PROGRAM ModeManagement_モード管理
VAR
    Setting_M : BOOL;
    Manual_M : BOOL;
    Auto_M : BOOL;
    Dummy_M : BOOL;
    Inital_M : BOOL;
    Output_Error_M : ARRAY[0..99] OF Bool;
    Index_Error_001 : DINT;
    Index_B_001 : DINT;
    Index_Share_001 : DINT;
    Error_TON : ARRAY[0..99] OF TON;  (* [2] A(左側) ST1 測定タイムアウト; [4] A(左側) ST5 測定タイムアウト *)
    Error_TOF : ARRAY[0..99] OF TOF;
    AutoMode_A_M : ARRAY[0..99] OF Bool;
    ６ : DINT;
    ST4_A_Rev_01_Origin_M : ARRAY[0..99] OF Bool;  (* A(左側) ST4 反転1 原点復帰工程; [1] A(左側) ST4 反転1 原点復帰開始; [2] A(左側) ST4 反転1 原点復帰中; [3] A(左側) ST4 反転1 ピックアップ戻; [4] A(左側) ST4 反転1 モータ原点復帰開始; [5] A(左側) ST4 反転1 ピックアップ行; [6] A(左側) ST4 反転1 チャック閉; [7] A(左側) ST4 反転1 原点復帰完了（ワーク無） *)
    ST4_A_Rev_01_OriginDone : BOOL;  (* A(左側) ST4 反転1 原点復帰完了 *)
    ST4_A_Rev_02_Origin_M : ARRAY[0..99] OF Bool;  (* A(左側) ST6 反転2 原点復帰工程; [1] A(左側) ST6 反転2 原点復帰開始; [2] A(左側) ST6 反転2 原点復帰中; [3] A(左側) ST6 反転2 ピックアップ戻; [4] A(左側) ST6 反転2 モータ原点復帰開始; [5] A(左側) ST6 反転2 ピックアップ行; [6] A(左側) ST6 反転2 チャック閉; [7] A(左側) ST6 反転2 原点復帰完了（ワーク無） *)
    ST4_A_Rev_02_OriginDone : BOOL;  (* A(左側) ST6 反転2 原点復帰完了 *)
    ST4_B_Rev_01_Origin_M : ARRAY[0..99] OF Bool;  (* B(右側) ST4 反転1 原点復帰工程; [1] B(右側) ST4 反転1 原点復帰開始; [2] B(右側) ST4 反転1 原点復帰中; [3] B(右側) ST4 反転1 ピックアップ戻; [4] B(右側) ST4 反転1 モータ原点復帰開始; [5] B(右側) ST4 反転1 ピックアップ行; [6] B(右側) ST4 反転1 チャック閉; [7] B(右側) ST4 反転1 原点復帰完了（ワーク無） *)
    ST4_B_Rev_01_OriginDone : BOOL;  (* B(右側) ST4 反転1 原点復帰完了 *)
    ST4_B_Rev_02_Origin_M : ARRAY[0..99] OF Bool;  (* B(右側) ST6 反転2 原点復帰工程; [1] B(右側) ST6 反転2 原点復帰開始; [2] B(右側) ST6 反転2 原点復帰中; [3] B(右側) ST6 反転2 ピックアップ戻; [4] B(右側) ST6 反転2 モータ原点復帰開始; [5] B(右側) ST6 反転2 ピックアップ行; [6] B(右側) ST6 反転2 チャック閉; [7] B(右側) ST6 反転2 原点復帰完了（ワーク無） *)
    ST4_B_Rev_02_OriginDone : BOOL;  (* B(右側) ST6 反転2 原点復帰完了 *)
END_VAR
VAR_EXTERNAL
    Output_A_Error_M : ARRAY[0..99] OF Bool;
    Output_A_Restart_M : ARRAY[0..99] OF Bool;
    In_Sw_RESET : BOOL;
    In_Sw_START : BOOL;
    ManualMode : BOOL;
    M9999 : BOOL;
    Output_B_Error_M : ARRAY[0..99] OF Bool;  (* B(右側)シリンダエラー *)
    Output_B_Restart_M : ARRAY[0..99] OF Bool;  (* B(右側)シリンダ再開： *)
    Output_Share_Error_M : ARRAY[0..99] OF Bool;
    Output_Share_Restart_M : ARRAY[0..99] OF Bool;
    TimerQ_In_Sen_Accum_CV_A_Full : BOOL;
    Out_TDC_Stop : BOOL;
    In_Sen_Unl_Conv_A_Pass : BOOL;
    In_Sen_Accum_CV_A_Full : BOOL;
    In_Sen_Unl_Conv_B_Pass : BOOL;
    Pause : ARRAY[0..99] OF Bool;  (* [3] FH A(左側) ST1; [9] FH A(左側) ST5; [10] FH B(右側) ST1; [11] FH B(右側) ST5; [12] A(左側) ST6 反転2 ワーク不一致 *)
    AutoMode : BOOL;
    In_Sen_DOOR_01 : BOOL;
    In_Sen_DOOR_02 : BOOL;
    In_Sen_DOOR_03 : BOOL;
    In_Sen_DOOR_04 : BOOL;
    In_Sen_DOOR_05 : BOOL;
    In_Sen_DOOR_06 : BOOL;
    In_Sw_EMS1 : BOOL;
    In_Sw_EMS2 : BOOL;
    In_Sw_EMS3 : BOOL;
    In_Sen_AIR１_Pressure_01 : BOOL;
    In_Sen_AIR１_Pressure_02 : BOOL;
    In_Sen_AIR１_Pressure_03 : BOOL;
    TEST_M : ARRAY[0..99] OF Bool;
    ST0_Sup_Start : BOOL;  (* ST0_動作開始 *)
    Out_CYw_Sply_Pick_A_H_Auto : ARRAY[0..10] OF Bool;
    Out_CYw_Sply_Pick_A_H_Done : BOOL;
    Out_CYw_Sply_Slide_A_H_Auto : ARRAY[0..10] OF Bool;
    Out_CYw_Sply_Slide_A_H_Done : BOOL;
    Out_CYw_Sup_Chuck_A_Cl_H_Auto : ARRAY[0..10] OF Bool;
    Out_CYw_Sup_Chuck_A_Cl_H_Done : BOOL;
    In_Sen_Accum_CV_A_Arrival : BOOL;
    In_Sen_Work_A_Pos_00 : BOOL;
    Out_CYw_Sply_Pick_A_F_Auto : ARRAY[0..10] OF Bool;
    Out_CYw_Sply_Pick_A_F_Done : BOOL;
    Out_CYw_Sup_Chuck_A_Cl_F_Auto : ARRAY[0..10] OF Bool;
    Out_CYw_Sup_Chuck_A_Cl_F_Done : BOOL;
    Out_CYw_Sply_Slide_A_F_Auto : ARRAY[0..10] OF Bool;
    Out_CYw_Sply_Slide_A_F_Done : BOOL;
    Ins_A_Cv_Error : BOOL;
    Station_A_Data : ARRAY[0..8] OF sData;
    Ins_A_Cv_M : ARRAY[0..99] OF Bool;
    HMI_MessageNo : ARRAY[0..9] OF UINT;
    FH_5552_10_A_Auto : BOOL;
    In_Sen_Accum_CV_B_Full : BOOL;
    FH_Line3_Error_Status_1 : BOOL;
    FH_Line0_Error_Status_1 : BOOL;
    FH_Line1_Error_Status_1 : BOOL;
    FH_Line2_Error_Status_1 : BOOL;
    FH_Line0_Error_Clear_1 : BOOL;
    FH_Line1_Error_Clear_1 : BOOL;
    FH_Line2_Error_Clear_1 : BOOL;
    FH_Line3_Error_Clear_1 : BOOL;
    Ins_A_Next_Cycle : BOOL;
    OriginDone : BOOL;  (* 原点復帰完了 *)
    DummyDone : BOOL;  (* ダミーチェック完了 *)
    HMI_CurrentPage : STRING[256];
    Ins_A_End : BOOL;
    Auto_A_Start : BOOL;  (* 自動運転 開始 *)
    Auto_Ready : BOOL;  (* 自動運転可能 *)
    ST0_A_Sup_Busy : BOOL;
    ST1_A_Ca1_Busy : BOOL;
    RCON1_1_IN_Alarm : BOOL;  (* 軸異常 *)
    RCON1_1_IN_EmergencyStop : BOOL;  (* 非常停止状態（監視） *)
    RCON1_1_Error : BOOL;  (* 異常予備（未接続） *)
    RCON1_1_IN_HomeDone : BOOL;  (* 原点復帰完了 *)
    RCON1_1_Error_Clear : BOOL;  (* 解除予備（未接続） *)
    Error_M : ARRAY[0..99] OF Bool;  (* エラー：; [1] シリンダ; [2] コンベア＆ドアセンサ; [3] FH A(左側) ST1; [4] A(左側)検査コンベア ワーク不一致; [5] RCON1-1 異常; [9] FH A(左側) ST5; [10] FH B(右側) ST1; [11] FH B(右側) ST5; [12] A(左側) ST6 反転2 ワーク不一致 *)
    ST1_A_Ca1_M : ARRAY[0..99] OF Bool;  (* [6] A(左側) ST1 検査前ワーク不一致 *)
    ST2_A_Hgt_M : ARRAY[0..99] OF Bool;
    ST3_A_Dis1_M : ARRAY[0..99] OF Bool;
    HMI_Home_SW : BOOL;
    Origin_Busy : BOOL;  (* 原点復帰中 *)
    Out_CYw_Rev_01_Pick_A_H_Origin : ARRAY[0..10] OF Bool;  (* 原点復帰【Y710】A(左側)ST4 反転1ピックアップ戻： *)
    Out_CYw_Rev_01_Pick_A_H_Done : BOOL;  (* 【Y710】A(左側)ST4 反転1ピックアップ戻 動作完了 *)
    Stm_A_Rev_Axis000_Origin : BOOL;  (* A(左側) ST4 反転1 モータ原点復帰開始 *)
    Stm_A_Rev_Axis000_OriginDone : BOOL;  (* A(左側) ST4 反転1 モータ原点復帰完了 *)
    Out_CYw_Rev_01_Pick_A_F_Origin : ARRAY[0..99] OF Bool;  (* 原点復帰【Y711】A(左側)ST4 反転1ピックアップ行： *)
    Out_CYw_Rev_01_Pick_A_F_Done : BOOL;  (* 【Y711】A(左側)ST4 反転1ピックアップ行 動作完了 *)
    Out_CYw_Rev_01_Chk_A_H_Origin : ARRAY[0..99] OF Bool;  (* 原点復帰【Y708】A(左側)ST4 反転1チャック閉： *)
    Out_CYw_Rev_01_Chk_A_H_Done : BOOL;  (* 【Y708】A(左側)ST4 反転1チャック閉 動作完了 *)
    TimerQ_In_Sen_Work_A_Pos_04 : BOOL;
    Out_CYw_Rev_02_Pick_A_H_Origin : ARRAY[0..10] OF Bool;  (* 原点復帰 【Y714】A(左側)ST6 反転2ピックアップ戻 *)
    Out_CYw_Rev_02_Pick_A_H_Done : BOOL;  (* 【Y714】A(左側)ST6 反転2ピックアップ戻 動作完了 *)
    Stm_A_Rev_Axis001_Origin : BOOL;  (* A(左側) ST6 反転2 モータ原点復帰開始 *)
    Stm_A_Rev_Axis001_OriginDone : BOOL;  (* A(左側) ST6 反転2 モータ原点復帰完了 *)
    Out_CYw_Rev_02_Pick_A_F_Origin : ARRAY[0..99] OF Bool;  (* 原点復帰 【Y715】A(左側)ST6 反転2ピックアップ行 *)
    Out_CYw_Rev_02_Pick_A_F_Done : BOOL;  (* 【Y715】A(左側)ST6 反転2ピックアップ行 動作完了 *)
    Out_CYw_Rev_02_Chk_A_H_Origin : ARRAY[0..99] OF Bool;  (* 原点復帰 【Y712】A(左側)ST6 反転2チャック閉 戻 *)
    Out_CYw_Rev_02_Chk_A_H_Done : BOOL;  (* 【Y712】A(左側)ST6 反転2チャック閉 戻 動作完了 *)
    TimerQ_In_Sen_Work_A_Pos_06 : BOOL;  (* 【X208】A(左側)ワーク位置6 *)
    Auto_B_Start : BOOL;  (* B(右側)自動運転開始（後続処理未接続） *)
    Out_CYw_Rev_01_Pick_B_H_Origin : ARRAY[0..10] OF Bool;  (* 原点復帰 【Y810】B(右側)ST4 反転1ピックアップ戻 *)
    Out_CYw_Rev_01_Pick_B_H_Done : BOOL;  (* 【Y810】B(右側)ST4 反転1ピックアップ戻 動作完了 *)
    Stm_B_Rev_Axis002_Origin : BOOL;  (* B(右側) ST4 反転1 モータ原点復帰開始 *)
    Stm_B_Rev_Axis002_OriginDone : BOOL;  (* B(右側) ST4 反転1 モータ原点復帰完了 *)
    Out_CYw_Rev_01_Pick_B_F_Origin : ARRAY[0..99] OF Bool;  (* 原点復帰 【Y811】B(右側)ST4 反転1ピックアップ行 *)
    Out_CYw_Rev_01_Pick_B_F_Done : BOOL;  (* 【Y811】B(右側)ST4 反転1ピックアップ行 動作完了 *)
    Out_CYw_Rev_01_Chk_B_H_Origin : ARRAY[0..99] OF Bool;  (* 原点復帰 【Y808】B(右側)ST4 反転1チャック閉 戻 *)
    Out_CYw_Rev_01_Chk_B_H_Done : BOOL;  (* 【Y808】B(右側)ST4 反転1チャック閉 戻 動作完了 *)
    TimerQ_In_Sen_Work_B_Pos_04 : BOOL;  (* 【X406】B(右側)ワーク位置4 *)
    Out_CYw_Rev_02_Pick_B_H_Origin : ARRAY[0..10] OF Bool;  (* 原点復帰 【Y814】B(右側)ST6 反転2ピックアップ戻 *)
    Out_CYw_Rev_02_Pick_B_H_Done : BOOL;  (* 【Y814】B(右側)ST6 反転2ピックアップ戻 動作完了 *)
    Stm_B_Rev_Axis003_Origin : BOOL;  (* B(右側) ST6 反転2 モータ原点復帰開始 *)
    Stm_B_Rev_Axis003_OriginDone : BOOL;  (* B(右側) ST6 反転2 モータ原点復帰完了 *)
    Out_CYw_Rev_02_Pick_B_F_Origin : ARRAY[0..99] OF Bool;  (* 原点復帰 【Y815】B(右側)ST6 反転2ピックアップ行 *)
    Out_CYw_Rev_02_Pick_B_F_Done : BOOL;  (* 【Y815】B(右側)ST6 反転2ピックアップ行 動作完了 *)
    Out_CYw_Rev_02_Chk_B_H_Origin : ARRAY[0..99] OF Bool;  (* 原点復帰 【Y812】B(右側)ST6 反転2チャック閉 戻 *)
    Out_CYw_Rev_02_Chk_B_H_Done : BOOL;  (* 【Y812】B(右側)ST6 反転2チャック閉 戻 動作完了 *)
    TimerQ_In_Sen_Work_B_Pos_06 : BOOL;  (* 【X408】B(右側)ワーク位置6 *)
    ST4_A_Rev1_M : ARRAY[0..99] OF Bool;  (* [10] A(左側) ST4 ワーク不一致エラー; [12] 【Y708】A(左側) ST4 反転1チャック閉 *)
    ST5_A_Ca2_M : ARRAY[0..99] OF Bool;  (* A(左側) ST5 カメラ2工程; [1] A(左側) ST5 カメラ2検査開始; [2] 【Y724】A(左側) ST5 ストッパー戻; [3] A(左側) ST5 ワーク有無判定; [4] A(左側) ST5 ワーク有; [5] A(左側) ST5 ワーク無; [6] A(左側) ST5 検査前ワーク不一致; [7] A(左側) ST5 FH測定開始 *)
    FH_A_ST5_Auto : BOOL;  (* A(左側) ST5 FH自動測定 *)
END_VAR
VAR_EXTERNAL CONSTANT
    ST6_A_Rev2_M : ARRAY[0..99] OF Bool;  (* A(左側) ST6 反転2工程; [1] A(左側) ST6 反転2 動作開始; [2] A(左側) ST6 反転2 【Y714】ピックアップ戻; [3] A(左側) ST6 反転2 【Y725】位置6ストッパー戻; [4] A(左側) ST6 反転2 原点角度転送; [5] A(左側) ST6 反転2 原点位置移動開始; [6] A(左側) ST6 反転2 原点位置移動完了; [7] A(左側) ST6 反転2 ワーク有無判定; [8] A(左側) ST6 反転2 ワーク有・前工程OK; [9] A(左側) ST6 反転2 ワーク無・前工程NG; [10] A(左側) ST6 反転2 ワーク不一致エラー; [11] A(左側) ST6 反転2 【Y715】反転前ピックアップ行; [12] A(左側) ST6 反転2 【Y712】チャック閉; [13] A(左側) ST6 反転2 【Y714】反転前ピックアップ戻; [14] A(左側) ST6 反転2 反転角度転送; [15] A(左側) ST6 反転2 反転位置移動完了; [16] A(左側) ST6 反転2 【Y715】設置ピックアップ行; [17] A(左側) ST6 反転2 【Y713】チャック開; [18] A(左側) ST6 反転2 【Y714】設置ピックアップ戻 *)
END_VAR
VAR_EXTERNAL
    ST7_A_Dis2_M : ARRAY[0..99] OF Bool;  (* [9] ST7 A ワーク有; [10] ST3 A ワーク無; [11] ST7 排出前ワーク不一致エラー; [12] コンベア下降 位置転送; [13] コンベア下降 移動開始; [14] 排出チャック開 行; [15] セイフティ上昇 位置転送; [16] セイフティ上昇 移動開始; [17] NG / フォルダストック 仕分け IAI移動位置 判定; [18] ストックフォルダ位置; [19] カメラ2 キズNG位置; [20] カメラ2 姿NG位置; [21] 排出フォルダ送り行; [22] SF/NG2左右 移動開始; [23] SF/NG2上下 目標位置転送; [24] ストックフォルダ カウントup; [25] カメラ キズNG位置; [26] カメラ 姿NG位置; [27] SF/NG2上下 移動開始; [28] 排出チャック戻／ワーク解放; [29] SF/NG2上下 原点位置転送; [30] SF/NG2上下 原点移動開始; [31] SF/NG2左右 原点位置転送; [32] 排出フォルダ送り戻; [33] 排出フォルダ戻完了 *)
END_VAR
VAR
    _p1 : BOOL;
    _p2 : BOOL;
    _p3 : BOOL;
    _p4 : BOOL;
    _p5 : BOOL;
    _p6 : BOOL;
    _p7 : BOOL;
    _p8 : BOOL;
    _p9 : BOOL;
    _p10 : BOOL;
    _p11 : BOOL;
    _p12 : BOOL;
    _p13 : BOOL;
    _p14 : BOOL;
    _p15 : BOOL;
    _p16 : BOOL;
    _p17 : BOOL;
    _p18 : BOOL;
    _p19 : BOOL;
    _p20 : BOOL;
    _p21 : BOOL;
    _p22 : BOOL;
    _p23 : BOOL;
    _p24 : BOOL;
    _e25 : R_TRIG;
    _e26 : R_TRIG;
    _e27 : R_TRIG;
    _e28 : R_TRIG;
    _e29 : R_TRIG;
    _e30 : R_TRIG;
    _e31 : R_TRIG;
    _e32 : R_TRIG;
    _e33 : R_TRIG;
    _p34 : BOOL;
    _p35 : BOOL;
    _p36 : BOOL;
    _p37 : BOOL;
    _p38 : BOOL;
    _p39 : BOOL;
    _p40 : BOOL;
    _e41 : R_TRIG;
    _p42 : BOOL;
    _e43 : R_TRIG;
    _e44 : R_TRIG;
    _e45 : R_TRIG;
    _e46 : R_TRIG;
    _e47 : R_TRIG;
    _e48 : R_TRIG;
    _e49 : R_TRIG;
    _p50 : BOOL;
    _p51 : BOOL;
    _p52 : BOOL;
    _p53 : BOOL;
    _p54 : BOOL;
    _p55 : BOOL;
    _p56 : BOOL;
END_VAR

(* Section Initial_初期化処理: ladder, written here as Structured Text *)

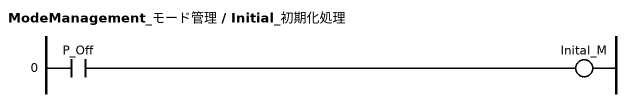
(* Rung 0 *)
Inital_M := P_Off;

(* Section Origin_原点復帰: ladder, written here as Structured Text *)

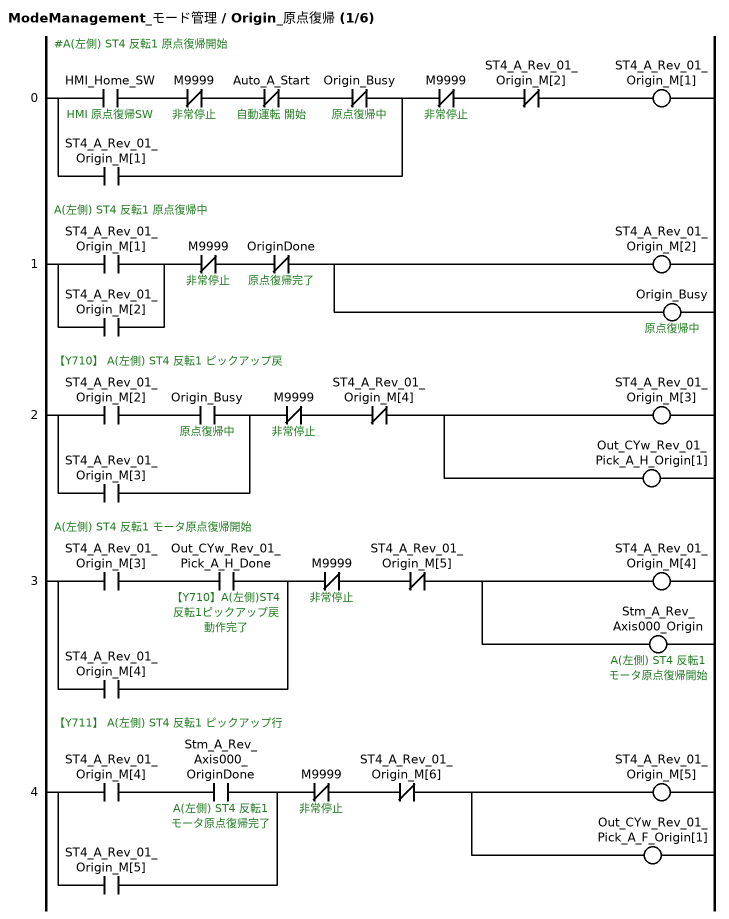
(* Rung 0: #A(左側) ST4 反転1 原点復帰開始 *)
ST4_A_Rev_01_Origin_M[1] := ((HMI_Home_SW AND NOT M9999 AND NOT Auto_A_Start AND NOT Origin_Busy) OR ST4_A_Rev_01_Origin_M[1]) AND NOT M9999 AND NOT ST4_A_Rev_01_Origin_M[2];
(* Rung 1: A(左側) ST4 反転1 原点復帰中 *)
_p1 := (ST4_A_Rev_01_Origin_M[1] OR ST4_A_Rev_01_Origin_M[2]) AND NOT M9999 AND NOT OriginDone;
ST4_A_Rev_01_Origin_M[2] := _p1;
Origin_Busy := _p1;
(* Rung 2: 【Y710】 A(左側) ST4 反転1 ピックアップ戻 *)
_p2 := ((ST4_A_Rev_01_Origin_M[2] AND Origin_Busy) OR ST4_A_Rev_01_Origin_M[3]) AND NOT M9999 AND NOT ST4_A_Rev_01_Origin_M[4];
ST4_A_Rev_01_Origin_M[3] := _p2;
Out_CYw_Rev_01_Pick_A_H_Origin[1] := _p2;
(* Rung 3: A(左側) ST4 反転1 モータ原点復帰開始 *)
_p3 := ((ST4_A_Rev_01_Origin_M[3] AND Out_CYw_Rev_01_Pick_A_H_Done) OR ST4_A_Rev_01_Origin_M[4]) AND NOT M9999 AND NOT ST4_A_Rev_01_Origin_M[5];
ST4_A_Rev_01_Origin_M[4] := _p3;
Stm_A_Rev_Axis000_Origin := _p3;
(* Rung 4: 【Y711】 A(左側) ST4 反転1 ピックアップ行 *)
_p4 := ((ST4_A_Rev_01_Origin_M[4] AND Stm_A_Rev_Axis000_OriginDone) OR ST4_A_Rev_01_Origin_M[5]) AND NOT M9999 AND NOT ST4_A_Rev_01_Origin_M[6];
ST4_A_Rev_01_Origin_M[5] := _p4;
Out_CYw_Rev_01_Pick_A_F_Origin[1] := _p4;

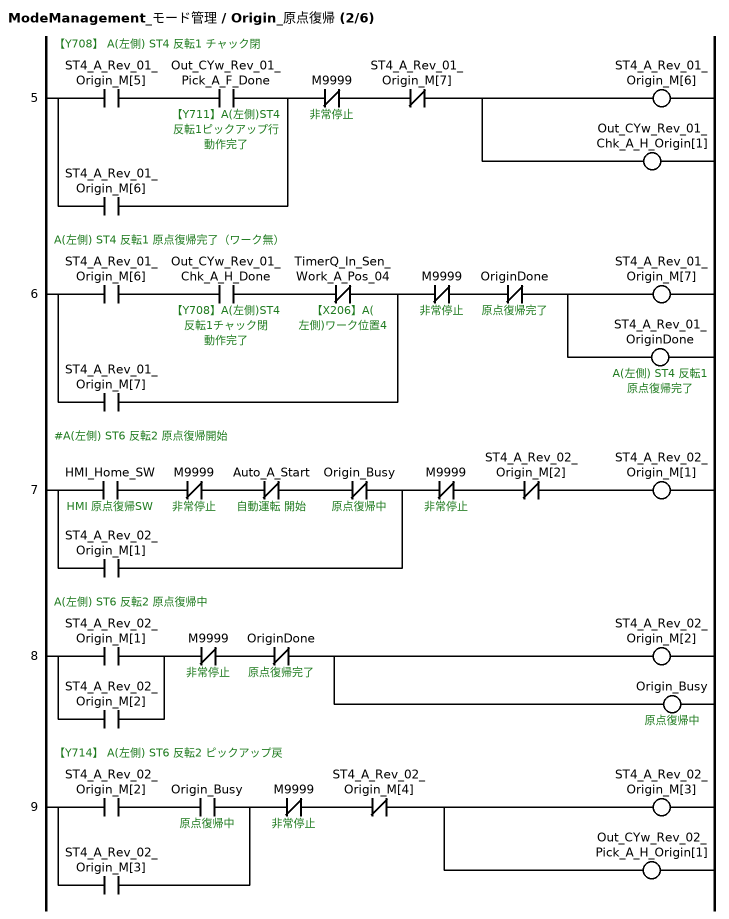
(* Rung 5: 【Y708】 A(左側) ST4 反転1 チャック閉 *)
_p5 := ((ST4_A_Rev_01_Origin_M[5] AND Out_CYw_Rev_01_Pick_A_F_Done) OR ST4_A_Rev_01_Origin_M[6]) AND NOT M9999 AND NOT ST4_A_Rev_01_Origin_M[7];
ST4_A_Rev_01_Origin_M[6] := _p5;
Out_CYw_Rev_01_Chk_A_H_Origin[1] := _p5;
(* Rung 6: A(左側) ST4 反転1 原点復帰完了（ワーク無） *)
_p6 := ((ST4_A_Rev_01_Origin_M[6] AND Out_CYw_Rev_01_Chk_A_H_Done AND NOT TimerQ_In_Sen_Work_A_Pos_04) OR ST4_A_Rev_01_Origin_M[7]) AND NOT M9999 AND NOT OriginDone;
ST4_A_Rev_01_Origin_M[7] := _p6;
ST4_A_Rev_01_OriginDone := _p6;
(* Rung 7: #A(左側) ST6 反転2 原点復帰開始 *)
ST4_A_Rev_02_Origin_M[1] := ((HMI_Home_SW AND NOT M9999 AND NOT Auto_A_Start AND NOT Origin_Busy) OR ST4_A_Rev_02_Origin_M[1]) AND NOT M9999 AND NOT ST4_A_Rev_02_Origin_M[2];
(* Rung 8: A(左側) ST6 反転2 原点復帰中 *)
_p7 := (ST4_A_Rev_02_Origin_M[1] OR ST4_A_Rev_02_Origin_M[2]) AND NOT M9999 AND NOT OriginDone;
ST4_A_Rev_02_Origin_M[2] := _p7;
Origin_Busy := _p7;
(* Rung 9: 【Y714】 A(左側) ST6 反転2 ピックアップ戻 *)
_p8 := ((ST4_A_Rev_02_Origin_M[2] AND Origin_Busy) OR ST4_A_Rev_02_Origin_M[3]) AND NOT M9999 AND NOT ST4_A_Rev_02_Origin_M[4];
ST4_A_Rev_02_Origin_M[3] := _p8;
Out_CYw_Rev_02_Pick_A_H_Origin[1] := _p8;

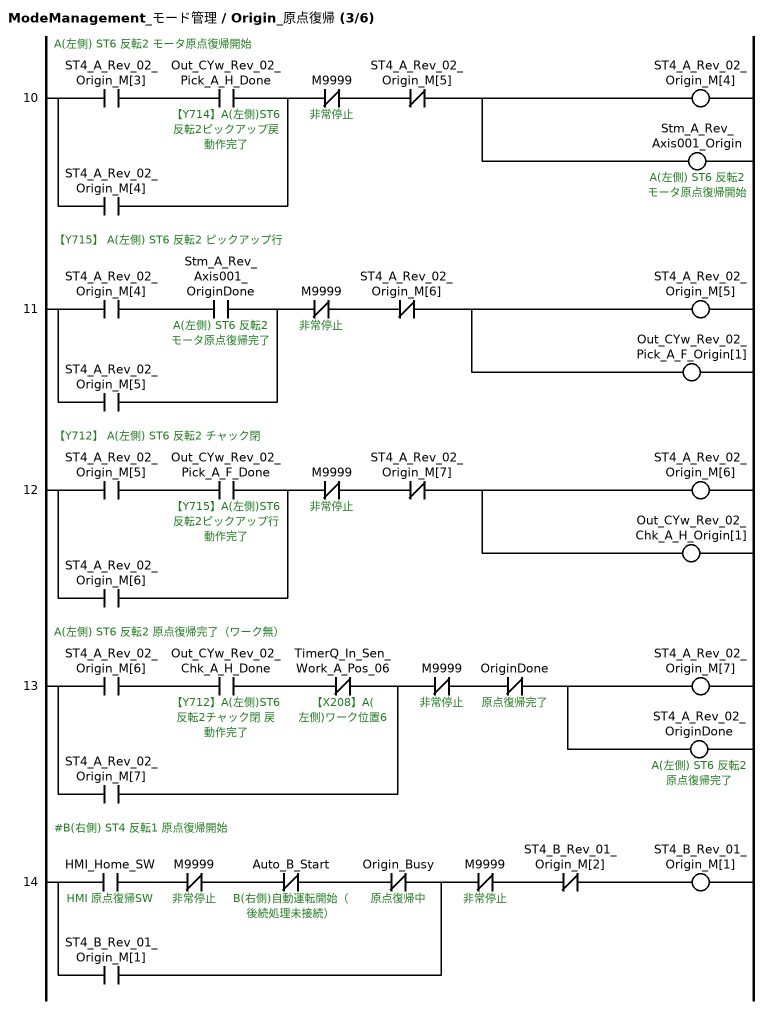
(* Rung 10: A(左側) ST6 反転2 モータ原点復帰開始 *)
_p9 := ((ST4_A_Rev_02_Origin_M[3] AND Out_CYw_Rev_02_Pick_A_H_Done) OR ST4_A_Rev_02_Origin_M[4]) AND NOT M9999 AND NOT ST4_A_Rev_02_Origin_M[5];
ST4_A_Rev_02_Origin_M[4] := _p9;
Stm_A_Rev_Axis001_Origin := _p9;
(* Rung 11: 【Y715】 A(左側) ST6 反転2 ピックアップ行 *)
_p10 := ((ST4_A_Rev_02_Origin_M[4] AND Stm_A_Rev_Axis001_OriginDone) OR ST4_A_Rev_02_Origin_M[5]) AND NOT M9999 AND NOT ST4_A_Rev_02_Origin_M[6];
ST4_A_Rev_02_Origin_M[5] := _p10;
Out_CYw_Rev_02_Pick_A_F_Origin[1] := _p10;
(* Rung 12: 【Y712】 A(左側) ST6 反転2 チャック閉 *)
_p11 := ((ST4_A_Rev_02_Origin_M[5] AND Out_CYw_Rev_02_Pick_A_F_Done) OR ST4_A_Rev_02_Origin_M[6]) AND NOT M9999 AND NOT ST4_A_Rev_02_Origin_M[7];
ST4_A_Rev_02_Origin_M[6] := _p11;
Out_CYw_Rev_02_Chk_A_H_Origin[1] := _p11;
(* Rung 13: A(左側) ST6 反転2 原点復帰完了（ワーク無） *)
_p12 := ((ST4_A_Rev_02_Origin_M[6] AND Out_CYw_Rev_02_Chk_A_H_Done AND NOT TimerQ_In_Sen_Work_A_Pos_06) OR ST4_A_Rev_02_Origin_M[7]) AND NOT M9999 AND NOT OriginDone;
ST4_A_Rev_02_Origin_M[7] := _p12;
ST4_A_Rev_02_OriginDone := _p12;
(* Rung 14: #B(右側) ST4 反転1 原点復帰開始 *)
ST4_B_Rev_01_Origin_M[1] := ((HMI_Home_SW AND NOT M9999 AND NOT Auto_B_Start AND NOT Origin_Busy) OR ST4_B_Rev_01_Origin_M[1]) AND NOT M9999 AND NOT ST4_B_Rev_01_Origin_M[2];

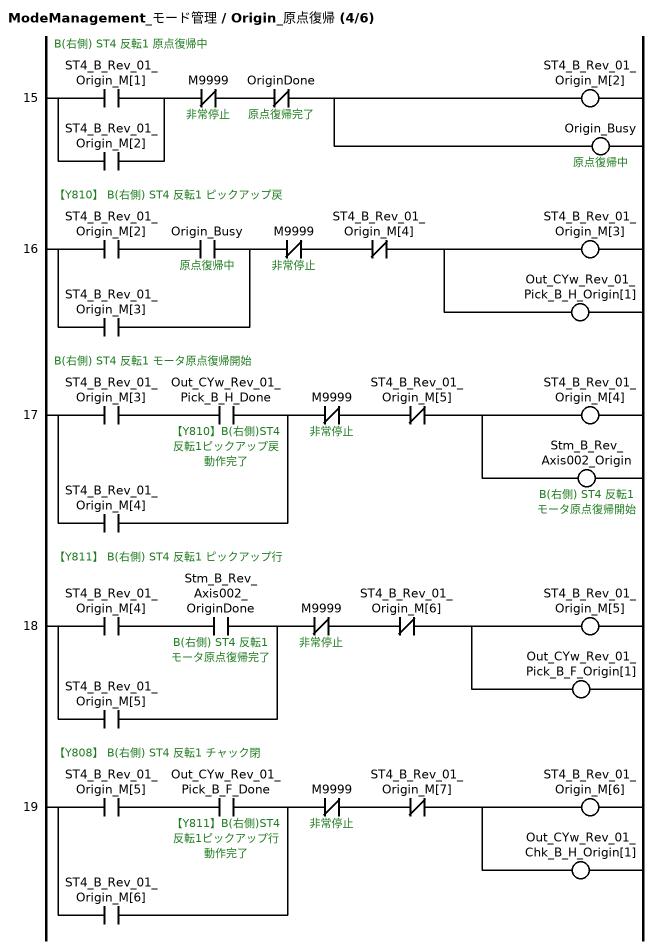
(* Rung 15: B(右側) ST4 反転1 原点復帰中 *)
_p13 := (ST4_B_Rev_01_Origin_M[1] OR ST4_B_Rev_01_Origin_M[2]) AND NOT M9999 AND NOT OriginDone;
ST4_B_Rev_01_Origin_M[2] := _p13;
Origin_Busy := _p13;
(* Rung 16: 【Y810】 B(右側) ST4 反転1 ピックアップ戻 *)
_p14 := ((ST4_B_Rev_01_Origin_M[2] AND Origin_Busy) OR ST4_B_Rev_01_Origin_M[3]) AND NOT M9999 AND NOT ST4_B_Rev_01_Origin_M[4];
ST4_B_Rev_01_Origin_M[3] := _p14;
Out_CYw_Rev_01_Pick_B_H_Origin[1] := _p14;
(* Rung 17: B(右側) ST4 反転1 モータ原点復帰開始 *)
_p15 := ((ST4_B_Rev_01_Origin_M[3] AND Out_CYw_Rev_01_Pick_B_H_Done) OR ST4_B_Rev_01_Origin_M[4]) AND NOT M9999 AND NOT ST4_B_Rev_01_Origin_M[5];
ST4_B_Rev_01_Origin_M[4] := _p15;
Stm_B_Rev_Axis002_Origin := _p15;
(* Rung 18: 【Y811】 B(右側) ST4 反転1 ピックアップ行 *)
_p16 := ((ST4_B_Rev_01_Origin_M[4] AND Stm_B_Rev_Axis002_OriginDone) OR ST4_B_Rev_01_Origin_M[5]) AND NOT M9999 AND NOT ST4_B_Rev_01_Origin_M[6];
ST4_B_Rev_01_Origin_M[5] := _p16;
Out_CYw_Rev_01_Pick_B_F_Origin[1] := _p16;
(* Rung 19: 【Y808】 B(右側) ST4 反転1 チャック閉 *)
_p17 := ((ST4_B_Rev_01_Origin_M[5] AND Out_CYw_Rev_01_Pick_B_F_Done) OR ST4_B_Rev_01_Origin_M[6]) AND NOT M9999 AND NOT ST4_B_Rev_01_Origin_M[7];
ST4_B_Rev_01_Origin_M[6] := _p17;
Out_CYw_Rev_01_Chk_B_H_Origin[1] := _p17;

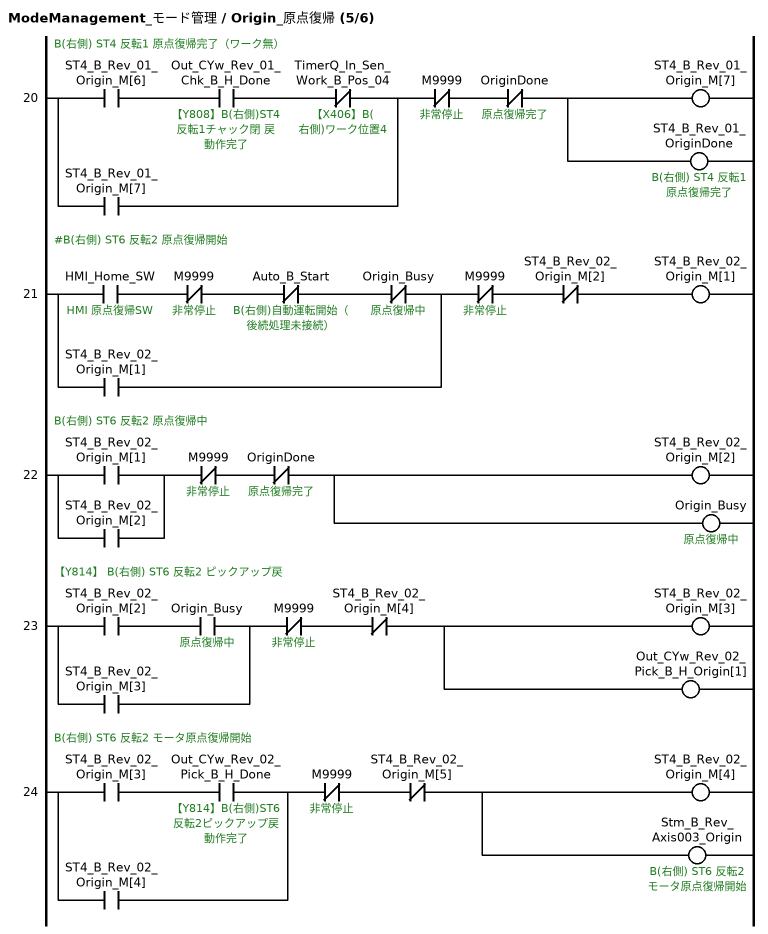
(* Rung 20: B(右側) ST4 反転1 原点復帰完了（ワーク無） *)
_p18 := ((ST4_B_Rev_01_Origin_M[6] AND Out_CYw_Rev_01_Chk_B_H_Done AND NOT TimerQ_In_Sen_Work_B_Pos_04) OR ST4_B_Rev_01_Origin_M[7]) AND NOT M9999 AND NOT OriginDone;
ST4_B_Rev_01_Origin_M[7] := _p18;
ST4_B_Rev_01_OriginDone := _p18;
(* Rung 21: #B(右側) ST6 反転2 原点復帰開始 *)
ST4_B_Rev_02_Origin_M[1] := ((HMI_Home_SW AND NOT M9999 AND NOT Auto_B_Start AND NOT Origin_Busy) OR ST4_B_Rev_02_Origin_M[1]) AND NOT M9999 AND NOT ST4_B_Rev_02_Origin_M[2];
(* Rung 22: B(右側) ST6 反転2 原点復帰中 *)
_p19 := (ST4_B_Rev_02_Origin_M[1] OR ST4_B_Rev_02_Origin_M[2]) AND NOT M9999 AND NOT OriginDone;
ST4_B_Rev_02_Origin_M[2] := _p19;
Origin_Busy := _p19;
(* Rung 23: 【Y814】 B(右側) ST6 反転2 ピックアップ戻 *)
_p20 := ((ST4_B_Rev_02_Origin_M[2] AND Origin_Busy) OR ST4_B_Rev_02_Origin_M[3]) AND NOT M9999 AND NOT ST4_B_Rev_02_Origin_M[4];
ST4_B_Rev_02_Origin_M[3] := _p20;
Out_CYw_Rev_02_Pick_B_H_Origin[1] := _p20;
(* Rung 24: B(右側) ST6 反転2 モータ原点復帰開始 *)
_p21 := ((ST4_B_Rev_02_Origin_M[3] AND Out_CYw_Rev_02_Pick_B_H_Done) OR ST4_B_Rev_02_Origin_M[4]) AND NOT M9999 AND NOT ST4_B_Rev_02_Origin_M[5];
ST4_B_Rev_02_Origin_M[4] := _p21;
Stm_B_Rev_Axis003_Origin := _p21;

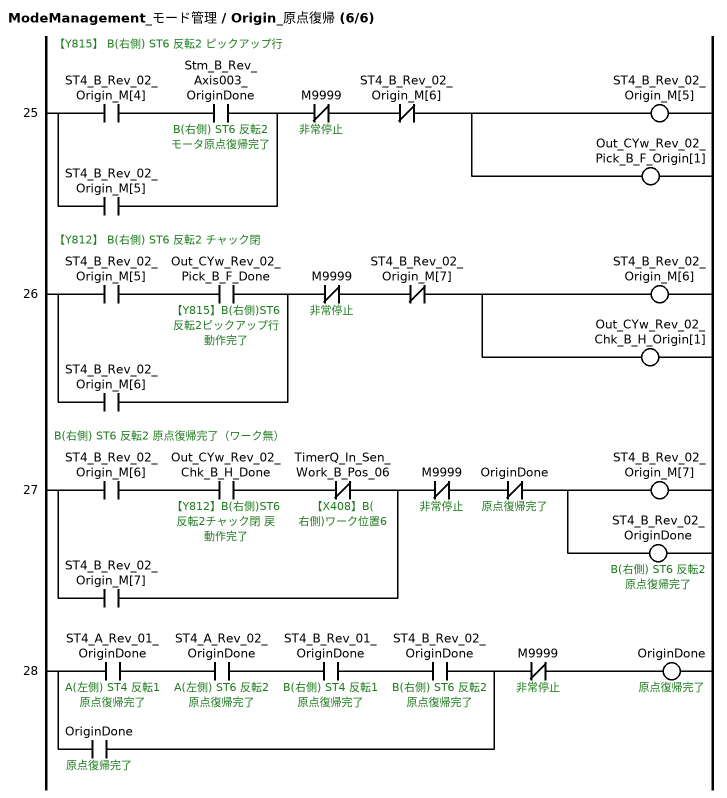
(* Rung 25: 【Y815】 B(右側) ST6 反転2 ピックアップ行 *)
_p22 := ((ST4_B_Rev_02_Origin_M[4] AND Stm_B_Rev_Axis003_OriginDone) OR ST4_B_Rev_02_Origin_M[5]) AND NOT M9999 AND NOT ST4_B_Rev_02_Origin_M[6];
ST4_B_Rev_02_Origin_M[5] := _p22;
Out_CYw_Rev_02_Pick_B_F_Origin[1] := _p22;
(* Rung 26: 【Y812】 B(右側) ST6 反転2 チャック閉 *)
_p23 := ((ST4_B_Rev_02_Origin_M[5] AND Out_CYw_Rev_02_Pick_B_F_Done) OR ST4_B_Rev_02_Origin_M[6]) AND NOT M9999 AND NOT ST4_B_Rev_02_Origin_M[7];
ST4_B_Rev_02_Origin_M[6] := _p23;
Out_CYw_Rev_02_Chk_B_H_Origin[1] := _p23;
(* Rung 27: B(右側) ST6 反転2 原点復帰完了（ワーク無） *)
_p24 := ((ST4_B_Rev_02_Origin_M[6] AND Out_CYw_Rev_02_Chk_B_H_Done AND NOT TimerQ_In_Sen_Work_B_Pos_06) OR ST4_B_Rev_02_Origin_M[7]) AND NOT M9999 AND NOT OriginDone;
ST4_B_Rev_02_Origin_M[7] := _p24;
ST4_B_Rev_02_OriginDone := _p24;
(* Rung 28 *)
OriginDone := ((ST4_A_Rev_01_OriginDone AND ST4_A_Rev_02_OriginDone AND ST4_B_Rev_01_OriginDone AND ST4_B_Rev_02_OriginDone) OR OriginDone) AND NOT M9999;

(* Section DummyCheck_ダミーチェック: ladder, written here as Structured Text *)

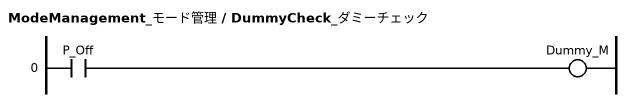
(* Rung 0 *)
Dummy_M := P_Off;

(* Section AutoMode_自動運転: ladder, written here as Structured Text *)

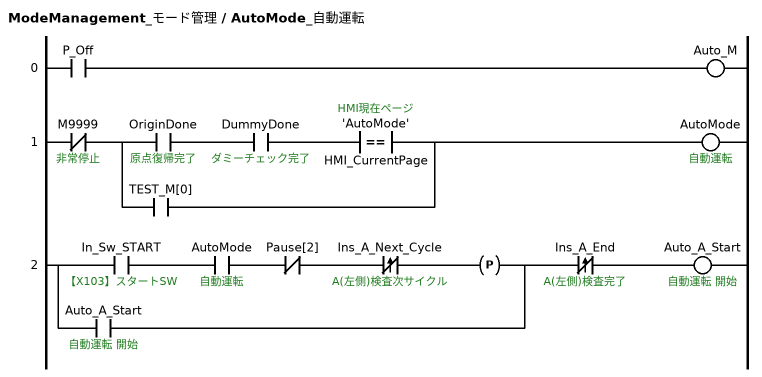
(* Rung 0 *)
Auto_M := P_Off;
(* Rung 1 *)
AutoMode := NOT M9999 AND ((OriginDone AND DummyDone AND ('AutoMode' = HMI_CurrentPage)) OR TEST_M[0]);
(* Rung 2 *)
_e25(CLK := Ins_A_Next_Cycle);
_e26(CLK := In_Sw_START AND AutoMode AND NOT Pause[2] AND NOT _e25.Q);
_e27(CLK := Ins_A_End);
Auto_A_Start := (_e26.Q OR Auto_A_Start) AND NOT _e27.Q;

(* Section Manual_手動運転: ladder, written here as Structured Text *)

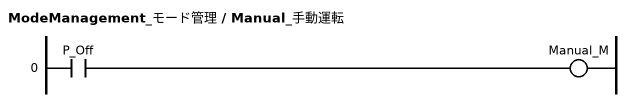
(* Rung 0 *)
Manual_M := P_Off;

(* Section Setting_設定: ladder, written here as Structured Text *)

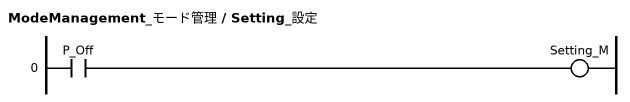
(* Rung 0 *)
Setting_M := P_Off;

(* Section Error_エラー処理: ladder, written here as Structured Text *)

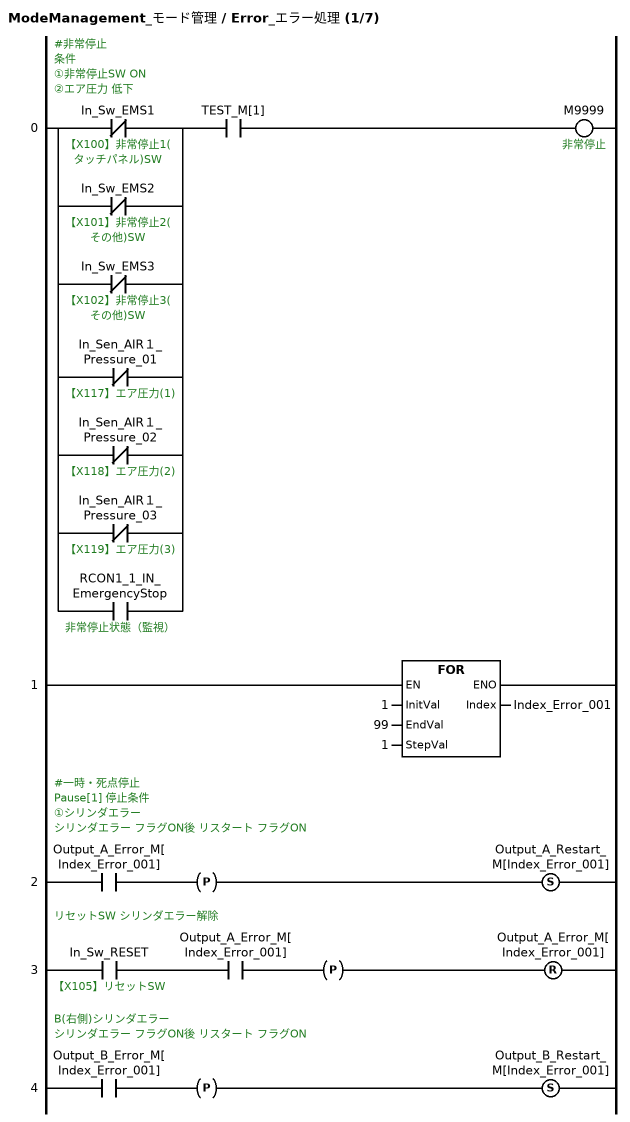
(* Rung 0: #非常停止 / 条件 / ①非常停止SW ON / ②エア圧力 低下 *)
M9999 := (NOT In_Sw_EMS1 OR NOT In_Sw_EMS2 OR NOT In_Sw_EMS3 OR NOT In_Sen_AIR１_Pressure_01 OR NOT In_Sen_AIR１_Pressure_02 OR NOT In_Sen_AIR１_Pressure_03 OR RCON1_1_IN_EmergencyStop) AND TEST_M[1];
(* Rung 1 *)
Index_Error_001 := FOR(InitVal := 1, EndVal := 99, StepVal := 1);
(* Rung 2: #一時・死点停止 / Pause[1] 停止条件 / ①シリンダエラー / シリンダエラー フラグON後 リスタート フラグON *)
_e28(CLK := Output_A_Error_M[Index_Error_001]);
IF _e28.Q THEN Output_A_Restart_M[Index_Error_001] := TRUE; END_IF;
(* Rung 3: リセットSW シリンダエラー解除 *)
_e29(CLK := In_Sw_RESET AND Output_A_Error_M[Index_Error_001]);
IF _e29.Q THEN Output_A_Error_M[Index_Error_001] := FALSE; END_IF;
(* Rung 4: B(右側)シリンダエラー / シリンダエラー フラグON後 リスタート フラグON *)
_e30(CLK := Output_B_Error_M[Index_Error_001]);
IF _e30.Q THEN Output_B_Restart_M[Index_Error_001] := TRUE; END_IF;

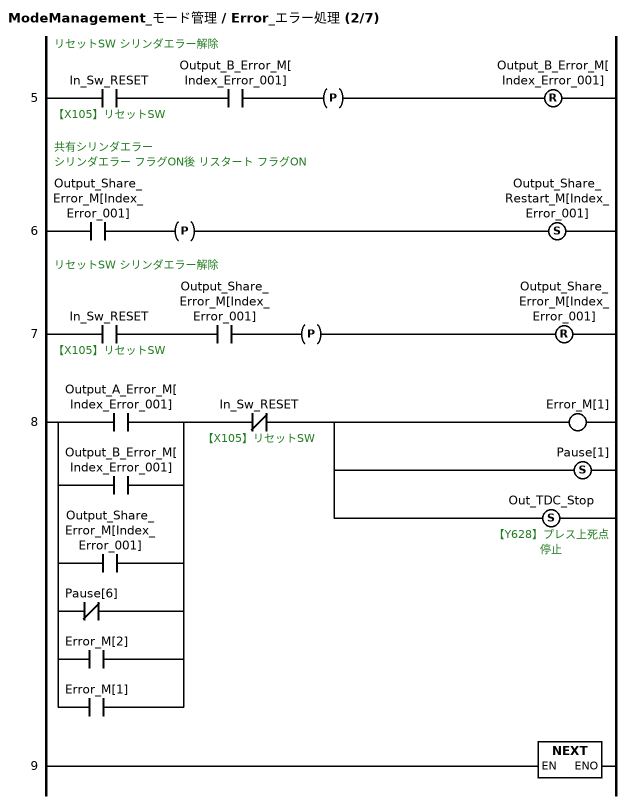
(* Rung 5: リセットSW シリンダエラー解除 *)
_e31(CLK := In_Sw_RESET AND Output_B_Error_M[Index_Error_001]);
IF _e31.Q THEN Output_B_Error_M[Index_Error_001] := FALSE; END_IF;
(* Rung 6: 共有シリンダエラー / シリンダエラー フラグON後 リスタート フラグON *)
_e32(CLK := Output_Share_Error_M[Index_Error_001]);
IF _e32.Q THEN Output_Share_Restart_M[Index_Error_001] := TRUE; END_IF;
(* Rung 7: リセットSW シリンダエラー解除 *)
_e33(CLK := In_Sw_RESET AND Output_Share_Error_M[Index_Error_001]);
IF _e33.Q THEN Output_Share_Error_M[Index_Error_001] := FALSE; END_IF;
(* Rung 8 *)
_p34 := (Output_A_Error_M[Index_Error_001] OR Output_B_Error_M[Index_Error_001] OR Output_Share_Error_M[Index_Error_001] OR NOT Pause[6] OR Error_M[2] OR Error_M[1]) AND NOT In_Sw_RESET;
Error_M[1] := _p34;
IF _p34 THEN
    Pause[1] := TRUE;
    Out_TDC_Stop := TRUE;
END_IF;
(* Rung 9 *)
NEXT();

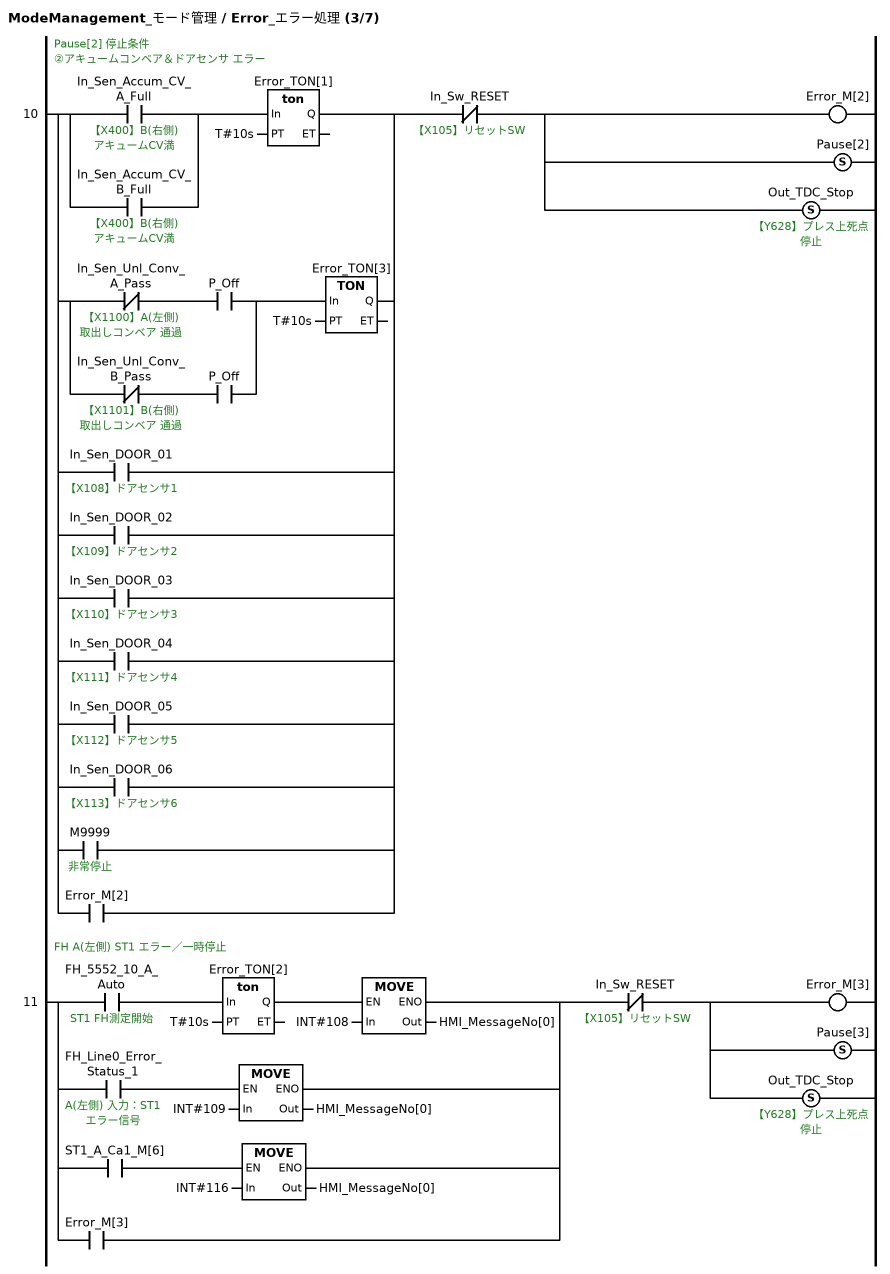
(* Rung 10: Pause[2] 停止条件 / ②アキュームコンベア＆ドアセンサ エラー *)
Error_TON[1](In := In_Sen_Accum_CV_A_Full OR In_Sen_Accum_CV_B_Full, PT := T#10s);
_p35 := Error_TON[1].Q;
Error_TON[3](In := (NOT In_Sen_Unl_Conv_A_Pass AND P_Off) OR (NOT In_Sen_Unl_Conv_B_Pass AND P_Off), PT := T#10s);
_p36 := (_p35 OR Error_TON[3].Q OR In_Sen_DOOR_01 OR In_Sen_DOOR_02 OR In_Sen_DOOR_03 OR In_Sen_DOOR_04 OR In_Sen_DOOR_05 OR In_Sen_DOOR_06 OR M9999 OR Error_M[2]) AND NOT In_Sw_RESET;
Error_M[2] := _p36;
IF _p36 THEN
    Pause[2] := TRUE;
    Out_TDC_Stop := TRUE;
END_IF;
(* Rung 11: FH A(左側) ST1 エラー／一時停止 *)
Error_TON[2](In := FH_5552_10_A_Auto, PT := T#10s);
IF Error_TON[2].Q THEN HMI_MessageNo[0] := INT#108; END_IF;
IF FH_Line0_Error_Status_1 THEN HMI_MessageNo[0] := INT#109; END_IF;
IF ST1_A_Ca1_M[6] THEN HMI_MessageNo[0] := INT#116; END_IF;
_p37 := (Error_TON[2].Q OR FH_Line0_Error_Status_1 OR ST1_A_Ca1_M[6] OR Error_M[3]) AND NOT In_Sw_RESET;
Error_M[3] := _p37;
IF _p37 THEN
    Pause[3] := TRUE;
    Out_TDC_Stop := TRUE;
END_IF;

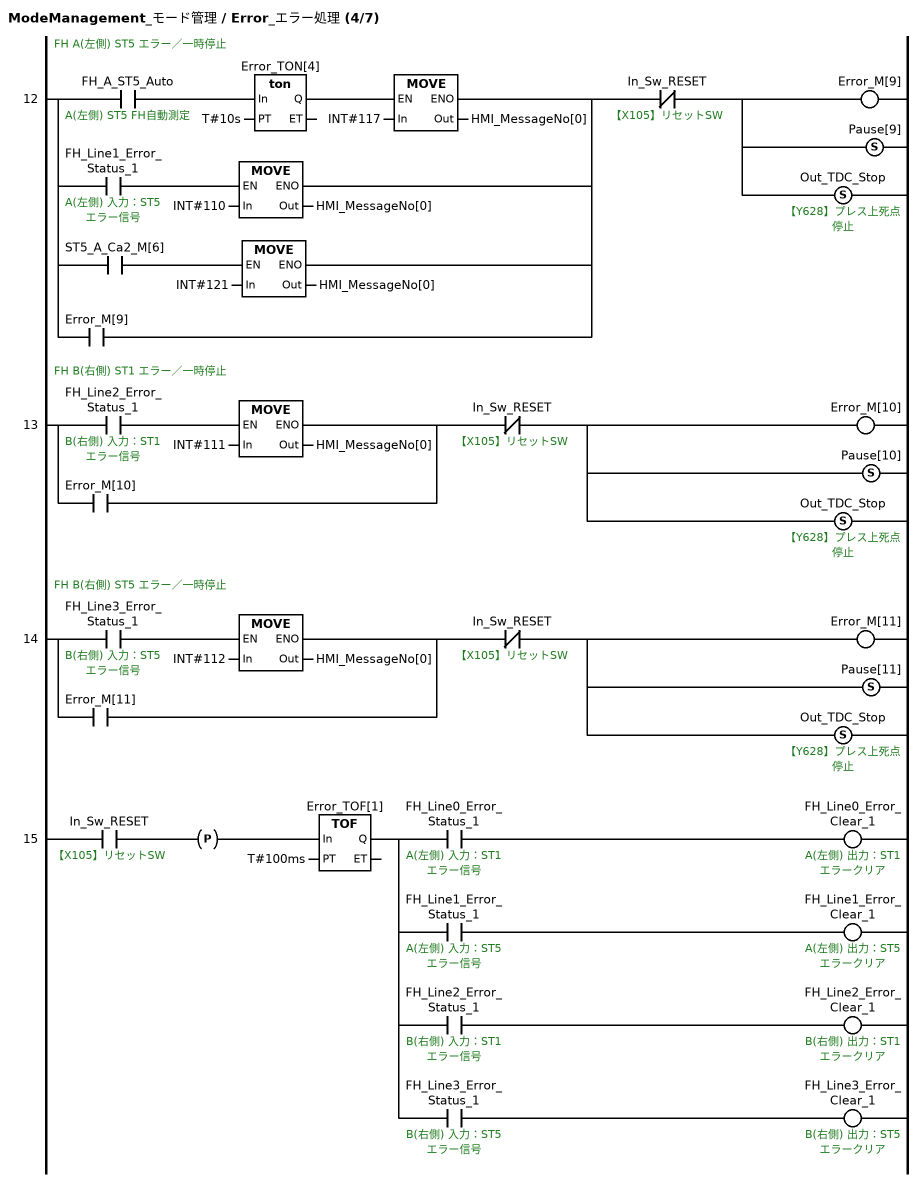
(* Rung 12: FH A(左側) ST5 エラー／一時停止 *)
Error_TON[4](In := FH_A_ST5_Auto, PT := T#10s);
IF Error_TON[4].Q THEN HMI_MessageNo[0] := INT#117; END_IF;
IF FH_Line1_Error_Status_1 THEN HMI_MessageNo[0] := INT#110; END_IF;
IF ST5_A_Ca2_M[6] THEN HMI_MessageNo[0] := INT#121; END_IF;
_p38 := (Error_TON[4].Q OR FH_Line1_Error_Status_1 OR ST5_A_Ca2_M[6] OR Error_M[9]) AND NOT In_Sw_RESET;
Error_M[9] := _p38;
IF _p38 THEN
    Pause[9] := TRUE;
    Out_TDC_Stop := TRUE;
END_IF;
(* Rung 13: FH B(右側) ST1 エラー／一時停止 *)
IF FH_Line2_Error_Status_1 THEN HMI_MessageNo[0] := INT#111; END_IF;
_p39 := (FH_Line2_Error_Status_1 OR Error_M[10]) AND NOT In_Sw_RESET;
Error_M[10] := _p39;
IF _p39 THEN
    Pause[10] := TRUE;
    Out_TDC_Stop := TRUE;
END_IF;
(* Rung 14: FH B(右側) ST5 エラー／一時停止 *)
IF FH_Line3_Error_Status_1 THEN HMI_MessageNo[0] := INT#112; END_IF;
_p40 := (FH_Line3_Error_Status_1 OR Error_M[11]) AND NOT In_Sw_RESET;
Error_M[11] := _p40;
IF _p40 THEN
    Pause[11] := TRUE;
    Out_TDC_Stop := TRUE;
END_IF;
(* Rung 15 *)
_e41(CLK := In_Sw_RESET);
Error_TOF[1](In := _e41.Q, PT := T#100ms);
FH_Line0_Error_Clear_1 := Error_TOF[1].Q AND FH_Line0_Error_Status_1;
FH_Line1_Error_Clear_1 := Error_TOF[1].Q AND FH_Line1_Error_Status_1;
FH_Line2_Error_Clear_1 := Error_TOF[1].Q AND FH_Line2_Error_Status_1;
FH_Line3_Error_Clear_1 := Error_TOF[1].Q AND FH_Line3_Error_Status_1;

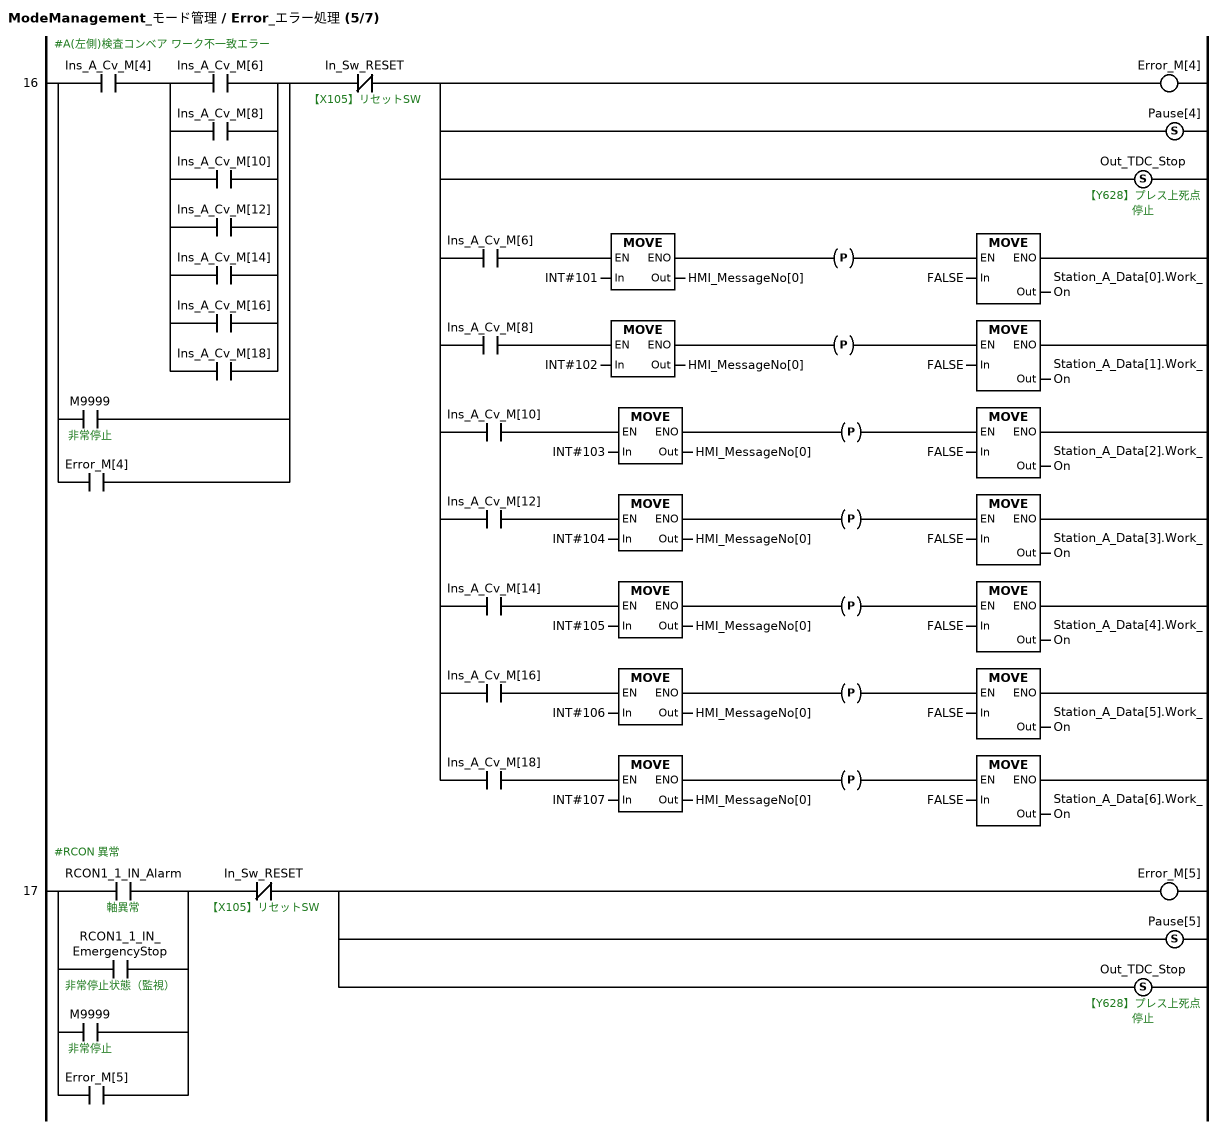
(* Rung 16: #A(左側)検査コンベア ワーク不一致エラー *)
_p42 := ((Ins_A_Cv_M[4] AND (Ins_A_Cv_M[6] OR Ins_A_Cv_M[8] OR Ins_A_Cv_M[10] OR Ins_A_Cv_M[12] OR Ins_A_Cv_M[14] OR Ins_A_Cv_M[16] OR Ins_A_Cv_M[18])) OR M9999 OR Error_M[4]) AND NOT In_Sw_RESET;
Error_M[4] := _p42;
IF _p42 THEN
    Pause[4] := TRUE;
    Out_TDC_Stop := TRUE;
END_IF;
IF _p42 AND Ins_A_Cv_M[6] THEN HMI_MessageNo[0] := INT#101; END_IF;
_e43(CLK := _p42 AND Ins_A_Cv_M[6]);
IF _e43.Q THEN Station_A_Data[0].Work_On := FALSE; END_IF;
IF _p42 AND Ins_A_Cv_M[8] THEN HMI_MessageNo[0] := INT#102; END_IF;
_e44(CLK := _p42 AND Ins_A_Cv_M[8]);
IF _e44.Q THEN Station_A_Data[1].Work_On := FALSE; END_IF;
IF _p42 AND Ins_A_Cv_M[10] THEN HMI_MessageNo[0] := INT#103; END_IF;
_e45(CLK := _p42 AND Ins_A_Cv_M[10]);
IF _e45.Q THEN Station_A_Data[2].Work_On := FALSE; END_IF;
IF _p42 AND Ins_A_Cv_M[12] THEN HMI_MessageNo[0] := INT#104; END_IF;
_e46(CLK := _p42 AND Ins_A_Cv_M[12]);
IF _e46.Q THEN Station_A_Data[3].Work_On := FALSE; END_IF;
IF _p42 AND Ins_A_Cv_M[14] THEN HMI_MessageNo[0] := INT#105; END_IF;
_e47(CLK := _p42 AND Ins_A_Cv_M[14]);
IF _e47.Q THEN Station_A_Data[4].Work_On := FALSE; END_IF;
IF _p42 AND Ins_A_Cv_M[16] THEN HMI_MessageNo[0] := INT#106; END_IF;
_e48(CLK := _p42 AND Ins_A_Cv_M[16]);
IF _e48.Q THEN Station_A_Data[5].Work_On := FALSE; END_IF;
IF _p42 AND Ins_A_Cv_M[18] THEN HMI_MessageNo[0] := INT#107; END_IF;
_e49(CLK := _p42 AND Ins_A_Cv_M[18]);
IF _e49.Q THEN Station_A_Data[6].Work_On := FALSE; END_IF;
(* Rung 17: #RCON 異常 *)
_p50 := (RCON1_1_IN_Alarm OR RCON1_1_IN_EmergencyStop OR M9999 OR Error_M[5]) AND NOT In_Sw_RESET;
Error_M[5] := _p50;
IF _p50 THEN
    Pause[5] := TRUE;
    Out_TDC_Stop := TRUE;
END_IF;

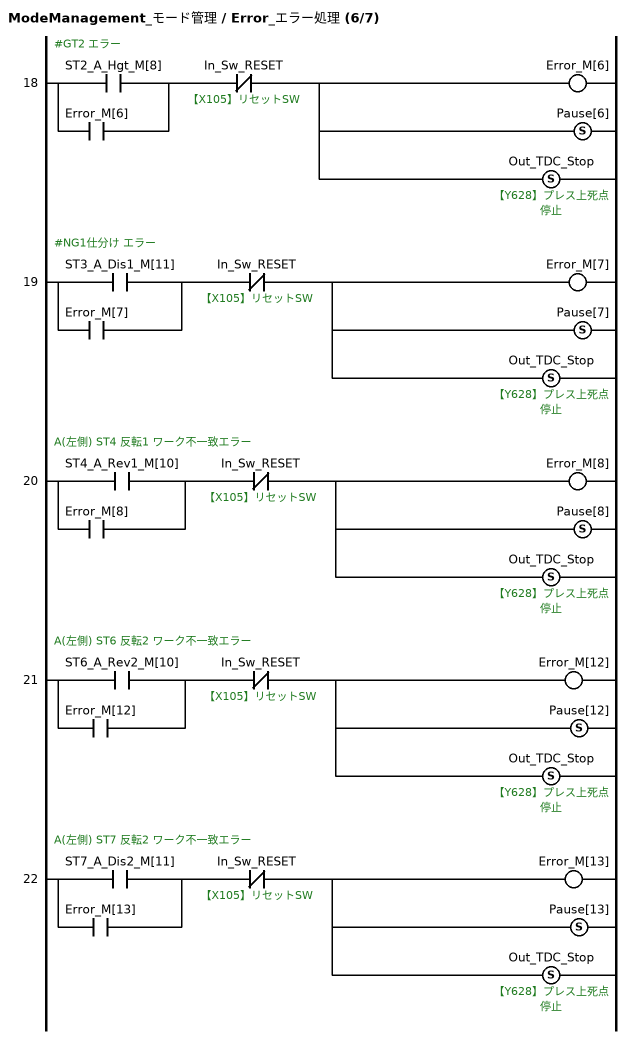
(* Rung 18: #GT2 エラー *)
_p51 := (ST2_A_Hgt_M[8] OR Error_M[6]) AND NOT In_Sw_RESET;
Error_M[6] := _p51;
IF _p51 THEN
    Pause[6] := TRUE;
    Out_TDC_Stop := TRUE;
END_IF;
(* Rung 19: #NG1仕分け エラー *)
_p52 := (ST3_A_Dis1_M[11] OR Error_M[7]) AND NOT In_Sw_RESET;
Error_M[7] := _p52;
IF _p52 THEN
    Pause[7] := TRUE;
    Out_TDC_Stop := TRUE;
END_IF;
(* Rung 20: A(左側) ST4 反転1 ワーク不一致エラー *)
_p53 := (ST4_A_Rev1_M[10] OR Error_M[8]) AND NOT In_Sw_RESET;
Error_M[8] := _p53;
IF _p53 THEN
    Pause[8] := TRUE;
    Out_TDC_Stop := TRUE;
END_IF;
(* Rung 21: A(左側) ST6 反転2 ワーク不一致エラー *)
_p54 := (ST6_A_Rev2_M[10] OR Error_M[12]) AND NOT In_Sw_RESET;
Error_M[12] := _p54;
IF _p54 THEN
    Pause[12] := TRUE;
    Out_TDC_Stop := TRUE;
END_IF;
(* Rung 22: A(左側) ST7 反転2 ワーク不一致エラー *)
_p55 := (ST7_A_Dis2_M[11] OR Error_M[13]) AND NOT In_Sw_RESET;
Error_M[13] := _p55;
IF _p55 THEN
    Pause[13] := TRUE;
    Out_TDC_Stop := TRUE;
END_IF;

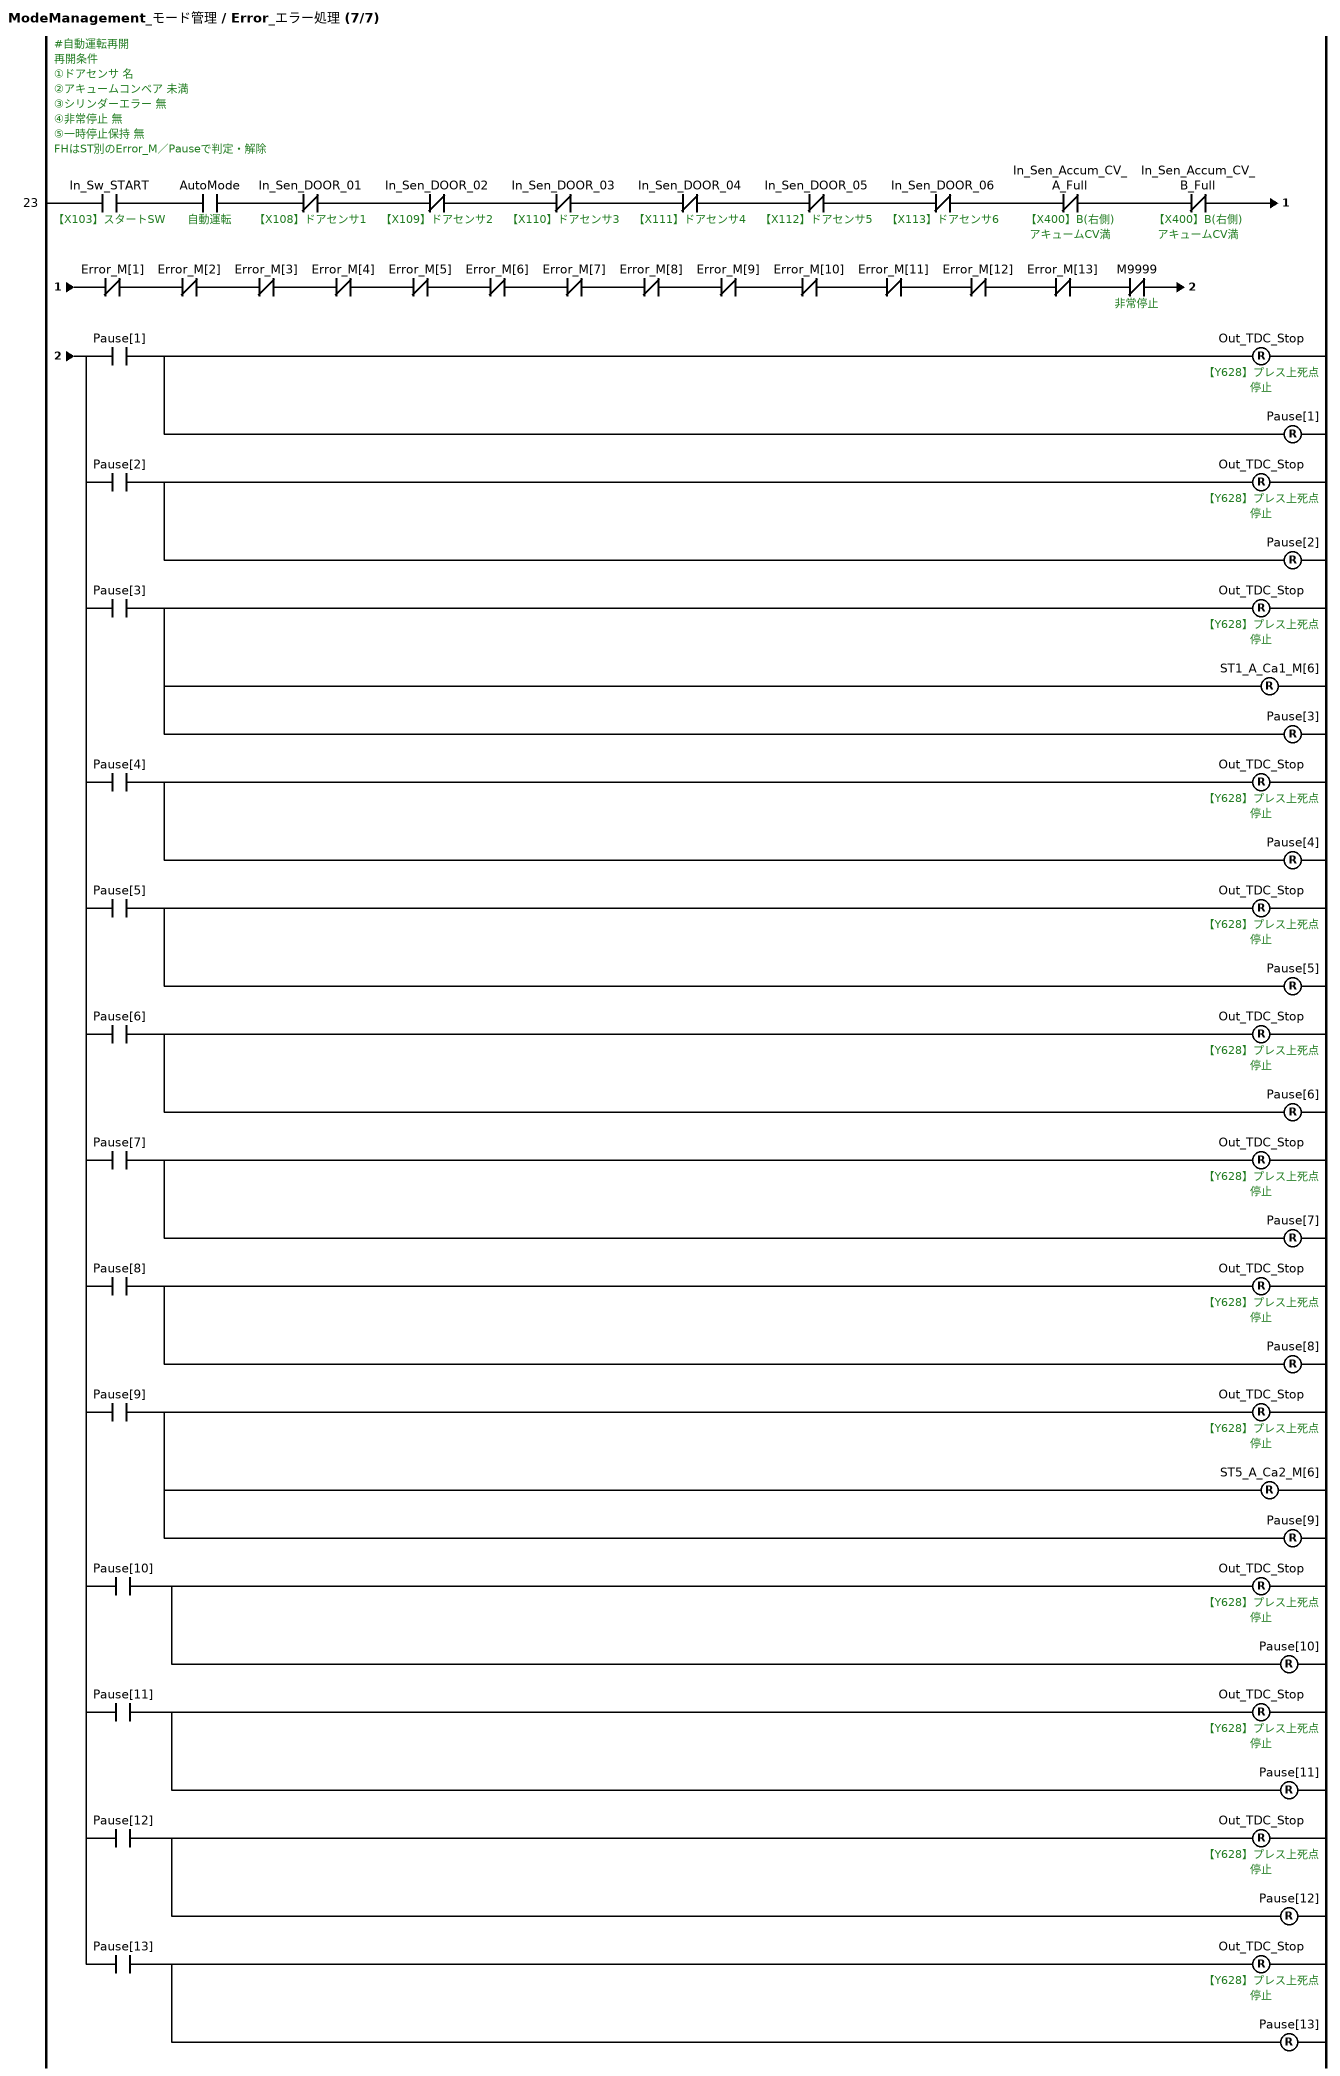
(* Rung 23: #自動運転再開 / 再開条件 / ①ドアセンサ 名 / ②アキュームコンベア 未満 / ③シリンダーエラー 無 / ④非常停止 無 / ⑤一時停止保持 無 / FHはST別のError_M／Pauseで判定・解除 *)
_p56 := In_Sw_START AND AutoMode AND NOT In_Sen_DOOR_01 AND NOT In_Sen_DOOR_02 AND NOT In_Sen_DOOR_03 AND NOT In_Sen_DOOR_04 AND NOT In_Sen_DOOR_05 AND NOT In_Sen_DOOR_06 AND NOT In_Sen_Accum_CV_A_Full AND NOT In_Sen_Accum_CV_B_Full AND NOT Error_M[1] AND NOT Error_M[2] AND NOT Error_M[3] AND NOT Error_M[4] AND NOT Error_M[5] AND NOT Error_M[6] AND NOT Error_M[7] AND NOT Error_M[8] AND NOT Error_M[9] AND NOT Error_M[10] AND NOT Error_M[11] AND NOT Error_M[12] AND NOT Error_M[13] AND NOT M9999;
IF _p56 AND Pause[1] THEN
    Out_TDC_Stop := FALSE;
    Pause[1] := FALSE;
END_IF;
IF _p56 AND Pause[2] THEN
    Out_TDC_Stop := FALSE;
    Pause[2] := FALSE;
END_IF;
IF _p56 AND Pause[3] THEN
    Out_TDC_Stop := FALSE;
    ST1_A_Ca1_M[6] := FALSE;
    Pause[3] := FALSE;
END_IF;
IF _p56 AND Pause[4] THEN
    Out_TDC_Stop := FALSE;
    Pause[4] := FALSE;
END_IF;
IF _p56 AND Pause[5] THEN
    Out_TDC_Stop := FALSE;
    Pause[5] := FALSE;
END_IF;
IF _p56 AND Pause[6] THEN
    Out_TDC_Stop := FALSE;
    Pause[6] := FALSE;
END_IF;
IF _p56 AND Pause[7] THEN
    Out_TDC_Stop := FALSE;
    Pause[7] := FALSE;
END_IF;
IF _p56 AND Pause[8] THEN
    Out_TDC_Stop := FALSE;
    Pause[8] := FALSE;
END_IF;
IF _p56 AND Pause[9] THEN
    Out_TDC_Stop := FALSE;
    ST5_A_Ca2_M[6] := FALSE;
    Pause[9] := FALSE;
END_IF;
IF _p56 AND Pause[10] THEN
    Out_TDC_Stop := FALSE;
    Pause[10] := FALSE;
END_IF;
IF _p56 AND Pause[11] THEN
    Out_TDC_Stop := FALSE;
    Pause[11] := FALSE;
END_IF;
IF _p56 AND Pause[12] THEN
    Out_TDC_Stop := FALSE;
    Pause[12] := FALSE;
END_IF;
IF _p56 AND Pause[13] THEN
    Out_TDC_Stop := FALSE;
    Pause[13] := FALSE;
END_IF;
END_PROGRAM

PROGRAM Movements_動作
VAR
    Mo_M : BOOL;
    ST0_A_Sup_M : ARRAY[0..99] OF Bool;  (* [4] 原点位置移動完了 *)
    ST1_Ins_Cv_Rdy : BOOL;
    ST2_Ins_Cv_Rdy : BOOL;
    ST3_Ins_Cv_Rdy : BOOL;
    ST4_Ins_Cv_Rdy : BOOL;
    ST5_Ins_Cv_Rdy : BOOL;
    ST6_Ins_Cv_Rdy : BOOL;
    ST7_Ins_Cv_Rdy : BOOL;
    Ins_A_Cv_T : ARRAY[0..99] OF TON;
    ST1_A_Ca1_Rdy : BOOL;
    GT2_A_Inspection_GetTime : DATE_AND_TIME;
    GT2_A_Inspection_GetTime_ST : STRING[256];
    GT2_A_Inspection_GetTime_ST_Del : STRING[20];
    ST4_A_Rev1_Busy : BOOL;  (* ST4 A 動作中 *)
    ST4_A_Rev_End : BOOL;
    ST6_A_Rev2_Busy : BOOL;  (* A(左側) ST6 反転2動作中 *)
    ST6_A_Rev2_End : BOOL;  (* A(左側) ST6 反転2動作完了 *)
    ST7_A_Dis2_Busy : BOOL;
    ST7_A_SF_M : ARRAY[0..99] OF Bool;
    ST7_A_SF_Busy : BOOL;
    ST7_A_SF_Wait_Pickup : BOOL;  (* フォルダストック取出し待ち *)
END_VAR
VAR_EXTERNAL
    ST0_Sup_Start : BOOL;  (* ST0_動作開始 *)
    M9999 : BOOL;
    Out_CYw_Sply_Pick_A_H_Auto : ARRAY[0..10] OF Bool;
    Out_CYw_Sply_Pick_A_H_Done : BOOL;
    Out_CYw_Sply_Slide_A_H_Auto : ARRAY[0..10] OF Bool;
    Out_CYw_Sply_Slide_A_H_Done : BOOL;
    Out_CYw_Sup_Chuck_A_Cl_H_Auto : ARRAY[0..10] OF Bool;
    Out_CYw_Sup_Chuck_A_Cl_H_Done : BOOL;
    In_Sen_Accum_CV_A_Arrival : BOOL;
    In_Sen_Work_A_Pos_00 : BOOL;
    Out_CYw_Sply_Pick_A_F_Auto : ARRAY[0..10] OF Bool;
    Out_CYw_Sply_Pick_A_F_Done : BOOL;
    Out_CYw_Sup_Chuck_A_Cl_F_Auto : ARRAY[0..10] OF Bool;
    Out_CYw_Sup_Chuck_A_Cl_F_Done : BOOL;
    Out_CYw_Sply_Slide_A_F_Auto : ARRAY[0..10] OF Bool;
    Out_CYw_Sply_Slide_A_F_Done : BOOL;
    Station_A_Data : ARRAY[0..8] OF sData;
    Cv_A_Data : ARRAY[0..8] OF sData;
    ST0_A_Sup_End : BOOL;  (* ST0 検査コンベア運転可 *)
    Out_CYS_Pos_01_Stopper_B_H_Auto : ARRAY[0..10] OF Bool;
    Out_CYS_Pos_02_Stopper_B_H_Auto : ARRAY[0..10] OF Bool;
    Out_CYS_Pos_03_Stopper_B_H_Auto : ARRAY[0..10] OF Bool;
    Out_CYS_Pos_04_Stopper_B_H_Auto : ARRAY[0..10] OF Bool;
    Out_CYS_Pos_05_Stopper_B_H_Auto : ARRAY[0..10] OF Bool;
    Out_CYS_Pos_06_Stopper_B_H_Auto : ARRAY[0..10] OF Bool;
    TimerQ_In_SenCY_Pos_01_Stopper_A_H : BOOL;
    TimerQ_In_SenCY_Pos_02_Stopper_A_H : BOOL;
    TimerQ_In_SenCY_Pos_03_Stopper_A_H : BOOL;
    TimerQ_In_SenCY_Pos_04_Stopper_A_H : BOOL;
    TimerQ_In_SenCY_Pos_05_Stopper_A_H : BOOL;
    TimerQ_In_SenCY_Pos_06_Stopper_A_H : BOOL;
    Out_Insp_Cv_A_Run_Auto : ARRAY[0..10] OF Bool;
    TimerQ_In_Sen_Work_A_Pos_01 : BOOL;
    TimerQ_In_Sen_Work_A_Pos_02 : BOOL;
    Pause : ARRAY[0..99] OF Bool;  (* [3] FH A(左側) ST1; [9] FH A(左側) ST5; [10] FH B(右側) ST1; [11] FH B(右側) ST5; [12] A(左側) ST6 反転2 ワーク不一致 *)
    TimerQ_In_Sen_Work_A_Pos_03 : BOOL;
    TimerQ_In_Sen_Work_A_Pos_04 : BOOL;
    TimerQ_In_Sen_Work_A_Pos_05 : BOOL;
    TimerQ_In_Sen_Work_A_Pos_06 : BOOL;
    TimerQ_In_Sen_Work_A_Pos_07 : BOOL;
    Out_CYS_Pos_01_Stopper_A_H_Auto : ARRAY[0..10] OF Bool;
    Out_CYS_Pos_02_Stopper_A_H_Auto : ARRAY[0..10] OF Bool;
    Out_CYS_Pos_03_Stopper_A_H_Auto : ARRAY[0..10] OF Bool;
    Out_CYS_Pos_04_Stopper_A_H_Auto : ARRAY[0..10] OF Bool;
    Out_CYS_Pos_05_Stopper_A_H_Auto : ARRAY[0..10] OF Bool;  (* [2] A(左側) ST5 カメラ2検査開始 *)
    Out_CYS_Pos_06_Stopper_A_H_Auto : ARRAY[0..10] OF Bool;  (* [1] A(左側)検査完了後; [2] A(左側) ST6 原点位置移動 *)
    Ins_A_Cv_M : ARRAY[0..99] OF Bool;
    Ins_A_Cv_Error : BOOL;  (* 検査コンベア ワーク不一致エラー *)
    TimerQ_In_Sen_Work_A_Pos_00 : BOOL;
    Out_CYS_Pos_01_Stopper_A_F_Auto : ARRAY[0..10] OF Bool;
    Out_CYS_Pos_02_Stopper_A_F_Auto : ARRAY[0..10] OF Bool;
    Out_CYS_Pos_03_Stopper_A_F_Auto : ARRAY[0..10] OF Bool;
    Out_CYS_Pos_04_Stopper_A_F_Auto : ARRAY[0..10] OF Bool;
    Out_CYS_Pos_05_Stopper_A_F_Auto : ARRAY[0..10] OF Bool;
    Out_CYS_Pos_06_Stopper_A_F_Auto : ARRAY[0..10] OF Bool;
    Ins_A_Next_Cycle : BOOL;  (* A(左側)検査コンベア 動作完了 *)
    ST0_A_Sup_Busy : BOOL;  (* ST0 稼働中 *)
    Ins_A_End : BOOL;  (* 検査完了 コンベア運転可能 *)
    Auto_A_Start : BOOL;
    Out_CYS_Pos_01_Stopper_A_H_Done : BOOL;
    FH_5552_10_A_Auto : BOOL;
    FH_A_ST1_Done : BOOL;
    ST1_A_Ca1_Busy : BOOL;  (* ST1 A検査中 *)
    ST1_A_Ca1_End : BOOL;  (* ST1 A 動作完了 *)
    ST2_A_Hgt_Busy : BOOL;  (* ST2 A 動作中 *)
    Out_CYw_HgtInsp_Clp_A_H_Auto : ARRAY[0..10] OF Bool;
    Out_CYw_HgtInsp_Clp_A_H_Done : BOOL;
    Out_CYw_HgtInsp_Lf_A_H_Auto : ARRAY[0..10] OF Bool;
    Out_CYw_HgtInsp_Lf_A_H_Done : BOOL;
    Out_CYS_Pos_02_Stopper_A_H_Done : BOOL;
    Out_CYw_HgtInsp_Clp_A_F_Auto : ARRAY[0..10] OF Bool;
    Out_CYw_HgtInsp_Clp_A_F_Done : BOOL;
    Out_CYw_HgtInsp_Lf_A_F_Auto : ARRAY[0..10] OF Bool;
    Out_CYw_HgtInsp_Lf_A_F_Done : BOOL;
    DLEP1_GT2_A_Auto : BOOL;
    Hgt_A_ComputedValueData : LREAL;
    Hight_LowerLimit : LREAL;  (* 高さ検査 下限値 *)
    Hight_UpperLimit : LREAL;  (* 高さ検査 上限値 *)
    ST2_A_Hgt_End : BOOL;  (* 高さ検査完了 *)
    ST3_A_Dis1_Busy : BOOL;  (* ST3 A 動作中 *)
    Out_CYw_NG1_Srt_A_H_Auto : ARRAY[0..10] OF Bool;
    Out_CYw_NG1_Srt_A_H_Done : BOOL;
    Out_CYw_Rev_01_Pick_A_H_Auto : ARRAY[0..10] OF Bool;  (* 自動【Y710】A(左側)ST4 反転1ピックアップ戻： *)
    Out_CYw_Rev_01_Pick_A_H_Done : BOOL;  (* 【Y710】A(左側)ST4 反転1ピックアップ戻 動作完了 *)
    Out_CYw_NG1_Pick_A_H_Auto : ARRAY[0..10] OF Bool;
    Out_CYw_NG1_Pick_A_H_Done : BOOL;
    Out_CYw_NG1_Chk_A_H_Auto : ARRAY[0..10] OF Bool;
    Out_CYw_NG1_Chk_A_H_Done : BOOL;
    RCON1_1_Auto : ARRAY[0..99] OF Bool;  (* 自動移動要求; [1] 原点位置移動; [2] NG仕分け; [3] 動作完了後 原点位置移動 *)
    RCON1_1_OUT_TargetPos_mm : LREAL;  (* 目標位置 [mm] *)
    HMI_RCON1_1_OUT_TargetPos : ARRAY[0..99] OF LREAL;  (* HMI設定位置 [mm]; [1] 原点位置; [3] 高さNG位置; [4] カメラ キズNG位置; [5] カメラ 姿NG位置 *)
    RCON1_1_M : ARRAY[0..99] OF BOOL;  (* #A(左側) RCON1_1 NG1排出(上下); [1] 開始指令保持; [2] 予備 *)
    RCON1_1_MoveDone : BOOL;  (* 動作完了 *)
    Error_M : ARRAY[0..99] OF Bool;  (* [3] FH A(左側) ST1; [9] FH A(左側) ST5; [10] FH B(右側) ST1; [11] FH B(右側) ST5; [12] A(左側) ST6 反転2 ワーク不一致 *)
    ST1_A_Ca1_M : ARRAY[0..99] OF Bool;  (* [1] ST1 A カメラ1 検査開始; [2] 【Y720】A(左側) 位置1ストッパー 戻; [3] ワーク有無 判定; [4] ST1 A ワーク有; [5] ST1 A ワーク無; [6] A(左側) ST1 検査前ワーク不一致; [7] ST1 FH測定開始 *)
    ST2_A_Hgt_M : ARRAY[0..99] OF Bool;  (* [4] 【Y721】A(左側) 位置2ストッパー戻; [6] ST1 A ワーク有; [7] ST1 A ワーク無; [5] ワーク有無 判定; [9] 【Y703】A(左側) 高さ検査持上行; [10] 【Y701】A(左側) 高さ検査押え行; [11] A(左側) 高さ検査OK判定; [12] A(左側) 高さ検査NG判定; [2] 【Y701】A(左側) 高さ検査押え行; [8] ST3 検査前ワーク不一致エラー *)
    Out_CYS_Pos_03_Stopper_A_H_Done : BOOL;
    Out_CYw_NG1_Pick_A_F_Auto : ARRAY[0..10] OF Bool;
    Out_CYw_NG1_Pick_A_F_Done : BOOL;
    Out_CYw_NG1_Chk_A_F_Auto : ARRAY[0..10] OF Bool;
    Out_CYw_NG1_Chk_A_F_Done : BOOL;
    Out_CYw_NG1_Srt_A_F_Auto : ARRAY[0..10] OF Bool;
    Out_CYw_NG1_Srt_A_F_Done : BOOL;
    ST3_A_Dis1_End : BOOL;  (* 左NG1排出 完了 *)
    ST3_A_Dis1_M : ARRAY[0..99] OF Bool;  (* [7] 原点位置 移動開始; [6] 原点位置移動 データ転送; [5] 【Y722】A(左側) 位置3ストッパー戻; [4] 【Y706】A(左側) NG1チャック戻; [8] ワーク有無 / 検査前ワーク不一致 判定; [9] S3 A ワーク有 工程NG; [10] S3 A ワーク無  前工程OK; [14] 【Y704】A(左側) NG1ピックアップ戻 ; [24] 仕分け完了 *)
    ST4_A_Rev1_M : ARRAY[0..99] OF Bool;  (* [2] ワーク有無 / 検査前ワーク不一致 判定; [3] 【Y723】A(左側) 位置4ストッパー戻; [4] ST4 A ワーク有; [5] ST4 A ワーク無 / 前工程NG; [6] ST4 検査前ワーク不一致エラー; [10] A(左側) ST4 ワーク不一致エラー; [12] 【Y708】A(左側) ST4 反転1チャック閉 *)
    Stm_A_Rev_Axis000_MovePos_Degree : LREAL;
    HMI_Stm_A_Rev_Axis000_MovePos_Degree : ARRAY[0..99] OF LREAL;  (* A(左側)ステッピングモータ000 回転角度 *)
    Stm_A_Rev_Axis000_Auto : ARRAY[0..99] OF Bool;  (* [1] 原点位置移動 開始 *)
    Stm_A_Rev_Axis000_MoveAbsoluteDone : BOOL;
    Out_CYw_Rev_01_Pick_A_F_Auto : ARRAY[0..10] OF Bool;
    Out_CYw_Rev_01_Pick_A_F_Done : BOOL;
    Out_CYw_Disc_Chk_A_H_Auto : ARRAY[0..10] OF Bool;
    Out_CYw_Disc_Chk_A_H_Done : BOOL;
    Out_CYw_Rev_02_Chk_A_H_Auto : ARRAY[0..10] OF Bool;
    Out_CYw_Rev_02_Chk_A_H_Done : BOOL;
    Out_CYw_Rev_02_Chk_A_F_Auto : ARRAY[0..10] OF Bool;
    Out_CYw_Rev_01_Chk_A_F_Auto : ARRAY[0..10] OF Bool;
    Out_CYw_Rev_01_Chk_A_F_Done : BOOL;
    ST5_A_Ca2_M : ARRAY[0..99] OF Bool;  (* A(左側) ST5 カメラ2工程; [1] A(左側) ST5 カメラ2検査開始; [2] 【Y724】A(左側) ST5 ストッパー戻; [3] A(左側) ST5 ワーク有無判定; [4] A(左側) ST5 ワーク有; [5] A(左側) ST5 ワーク無; [6] A(左側) ST5 検査前ワーク不一致; [7] A(左側) ST5 FH測定開始 *)
    ST5_A_Ca2_Busy : BOOL;  (* A(左側) ST5 カメラ2検査中 *)
    ST5_A_Ca2_End : BOOL;  (* A(左側) ST5 カメラ2動作完了 *)
    FH_A_ST5_Auto : BOOL;  (* A(左側) ST5 FH自動測定 *)
    FH_A_ST5_Done : BOOL;  (* A(左側) ST5 画像検査完了 *)
    Out_CYS_Pos_05_Stopper_A_H_Done : BOOL;  (* 【Y724】A(左側) 位置5ストッパー戻 動作完了 *)
    Out_CYw_Rev_01_Chk_A_H_Auto : ARRAY[0..10] OF Bool;  (* 自動【Y708】A(左側)ST4 反転1チャック閉： *)
    Out_CYw_Rev_01_Chk_A_H_Done : BOOL;  (* 【Y708】A(左側)ST4 反転1チャック閉 動作完了 *)
    HMI_Stm_A_Rev_Axis001_MovePos_Degree : ARRAY[0..99] OF LREAL;  (* A(左側) ST6 反転2設定角度; [1] A(左側) ST6 原点位置設定角度; [2] A(左側) ST6 反転位置設定角度 *)
    Out_CYw_Rev_02_Chk_A_F_Done : BOOL;  (* 【Y713】A(左側)ST6 反転2チャック開 行 動作完了 *)
    Out_CYw_Rev_02_Pick_A_F_Auto : ARRAY[0..10] OF Bool;  (* 自動【Y715】A(左側)ST6 反転2ピックアップ行 ：; [1] A(左側) ST6 反転前行; [2] A(左側) ST6 設置行 *)
    Out_CYw_Rev_02_Pick_A_F_Done : BOOL;  (* 【Y715】A(左側)ST6 反転2ピックアップ行 動作完了 *)
    Out_CYw_Rev_02_Pick_A_H_Auto : ARRAY[0..10] OF Bool;  (* 自動【Y714】A(左側)ST6 反転2ピックアップ戻 ：; [1] A(左側) ST6 反転前戻; [2] A(左側) ST6 設置後戻 *)
    Out_CYw_Rev_02_Pick_A_H_Done : BOOL;  (* 【Y714】A(左側)ST6 反転2ピックアップ戻 動作完了 *)
    Stm_A_Rev_Axis001_Auto : ARRAY[0..99] OF Bool;  (* A(左側) ST6 反転2自動指令; [1] A(左側) ST6 原点位置移動開始 *)
    Stm_A_Rev_Axis001_MoveAbsoluteDone : BOOL;  (* A(左側) ST6 反転2位置決め完了 *)
    Stm_A_Rev_Axis001_MovePos_Degree : LREAL;  (* A(左側) ST6 反転2指令角度 *)
    ST6_A_Rev2_M : ARRAY[0..99] OF Bool;
    RCON1_5_Auto : ARRAY[0..99] OF Bool;  (* 自動移動要求; [1] 原点位置移動; [2] 自動要求2（外部接続用）; [3] 自動要求3（外部接続用） *)
    HMI_RCON1_5_OUT_TargetPos : ARRAY[0..99] OF LREAL;  (* RCON1_5 目標位置 [mm]： *)
    RCON1_5_MoveDone : BOOL;
    Out_CYw_Ejc_Hldr_Feed_A_H_Auto : ARRAY[0..10] OF Bool;
    Out_CYw_Ejc_Hldr_Feed_A_H_Done : BOOL;
    HMI_RCON1_3_OUT_TargetPos : ARRAY[0..99] OF LREAL;  (* RCON1_3 SF/NG2仕分け(左右) 目標位置 [mm]： *)
    RCON1_3_Auto : ARRAY[0..99] OF Bool;
    RCON1_3_MoveDone : BOOL;
    ST7_A_Dis2_M : ARRAY[0..99] OF Bool;  (* [9] ST7 A ワーク有; [10] ST3 A ワーク無; [11] ST7 排出前ワーク不一致エラー; [12] コンベア下降 位置転送; [13] コンベア下降 移動開始; [14] 排出チャック開 行; [15] セイフティ上昇 位置転送; [16] セイフティ上昇 移動開始; [17] NG / フォルダストック 仕分け IAI移動位置 判定; [18] ストックフォルダ位置; [19] カメラ2 キズNG位置; [20] カメラ2 姿NG位置; [21] 排出フォルダ送り行; [22] SF/NG2左右 移動開始; [23] SF/NG2上下 目標位置転送; [24] ストックフォルダ カウントup; [25] カメラ キズNG位置; [26] カメラ 姿NG位置; [27] SF/NG2上下 移動開始; [28] 排出チャック戻／ワーク解放; [29] SF/NG2上下 原点位置転送; [30] SF/NG2上下 原点移動開始; [31] SF/NG2左右 原点位置転送; [32] 排出フォルダ送り戻; [33] 排出フォルダ戻完了 *)
    RCON1_3_OUT_TargetPos_mm : LREAL;
    A_SF_CT : INT;  (* A(左側) ストックフォルダカウント *)
    TimerQ_In_Sen_SH_B_Ent : BOOL;
    TimerQ_In_Sen_SH_B_Ext : BOOL;
    RCON1_5_ActualPos_mm : LREAL;
    RCON1_5_SafePos_mm : LREAL;
    Out_CYw_SH_A_Turn_F_Auto : ARRAY[0..10] OF Bool;
    TimerQ_In_SenCY_SH_A_Turn_F : BOOL;
    Out_CYw_SH_A_Turn_H_Auto : ARRAY[0..10] OF Bool;
    TimerQ_In_SenCY_SH_A_Turn_H : BOOL;
    Out_CYw_SH_A_Turn_H_Done : BOOL;
    Out_CYw_SH_A_Turn_F_Done : BOOL;
    Out_CYw_Ejc_Hldr_Feed_A_F_Auto : ARRAY[0..10] OF Bool;
    Out_CYw_Ejc_Hldr_Feed_A_F_Done : BOOL;
    Out_CYw_Disc_Chk_A_F_Auto : ARRAY[0..10] OF Bool;
    Out_CYw_Disc_Chk_A_F_Done : BOOL;
    RCON1_5_OUT_TargetPos_mm : LREAL;
END_VAR
VAR
    _e1 : R_TRIG;
    _p2 : BOOL;
    _e3 : R_TRIG;
    _e4 : R_TRIG;
    _p5 : BOOL;
    _e6 : R_TRIG;
    _e7 : R_TRIG;
    _p8 : BOOL;
    _p9 : BOOL;
    _p10 : BOOL;
    _p11 : BOOL;
    _p12 : BOOL;
    _p13 : BOOL;
    _p14 : BOOL;
    _p15 : BOOL;
    _e16 : R_TRIG;
    _p17 : BOOL;
    _p18 : BOOL;
    _p19 : BOOL;
    _p20 : BOOL;
    _p21 : BOOL;
    _p22 : BOOL;
    _p23 : BOOL;
    _p24 : BOOL;
    _p25 : BOOL;
    _p26 : BOOL;
    _p27 : BOOL;
    _p28 : BOOL;
    _e29 : R_TRIG;
    _p30 : BOOL;
    _e31 : R_TRIG;
    _p32 : BOOL;
    _p33 : BOOL;
    _p34 : BOOL;
    _p35 : BOOL;
    _p36 : BOOL;
    _e37 : R_TRIG;
    _p38 : BOOL;
    _p39 : BOOL;
    _p40 : BOOL;
    _p41 : BOOL;
    _p42 : BOOL;
    _p43 : BOOL;
    _p44 : BOOL;
    _p45 : BOOL;
    _p46 : BOOL;
    _e47 : R_TRIG;
    _p48 : BOOL;
    _p49 : BOOL;
    _p50 : BOOL;
    _p51 : BOOL;
    _p52 : BOOL;
    _p53 : BOOL;
    _p54 : BOOL;
    _p55 : BOOL;
    _p56 : BOOL;
    _p57 : BOOL;
    _p58 : BOOL;
    _p59 : BOOL;
    _p60 : BOOL;
    _p61 : BOOL;
    _e62 : R_TRIG;
    _p63 : BOOL;
    _p64 : BOOL;
    _p65 : BOOL;
    _p66 : BOOL;
    _p67 : BOOL;
    _p68 : BOOL;
    _p69 : BOOL;
    _p70 : BOOL;
    _e71 : R_TRIG;
    _p72 : BOOL;
    _p73 : BOOL;
    _p74 : BOOL;
    _p75 : BOOL;
    _p76 : BOOL;
    _e77 : R_TRIG;
    _p78 : BOOL;
    _p79 : BOOL;
    _p80 : BOOL;
    _p81 : BOOL;
    _p82 : BOOL;
    _p83 : BOOL;
    _p84 : BOOL;
    _p85 : BOOL;
    _p86 : BOOL;
    _p87 : BOOL;
    _p88 : BOOL;
    _e89 : R_TRIG;
    _p90 : BOOL;
    _p91 : BOOL;
    _p92 : BOOL;
    _p93 : BOOL;
    _p94 : BOOL;
    _e95 : R_TRIG;
    _p96 : BOOL;
    _p97 : BOOL;
    _p98 : BOOL;
    _p99 : BOOL;
    _p100 : BOOL;
    _p101 : BOOL;
    _p102 : BOOL;
    _e103 : R_TRIG;
    _p104 : BOOL;
    _p105 : BOOL;
    _e106 : R_TRIG;
    _p107 : BOOL;
    _p108 : BOOL;
    _p109 : BOOL;
END_VAR

(* Section Ins_A_Cv_左検査Cv: ladder, written here as Structured Text *)

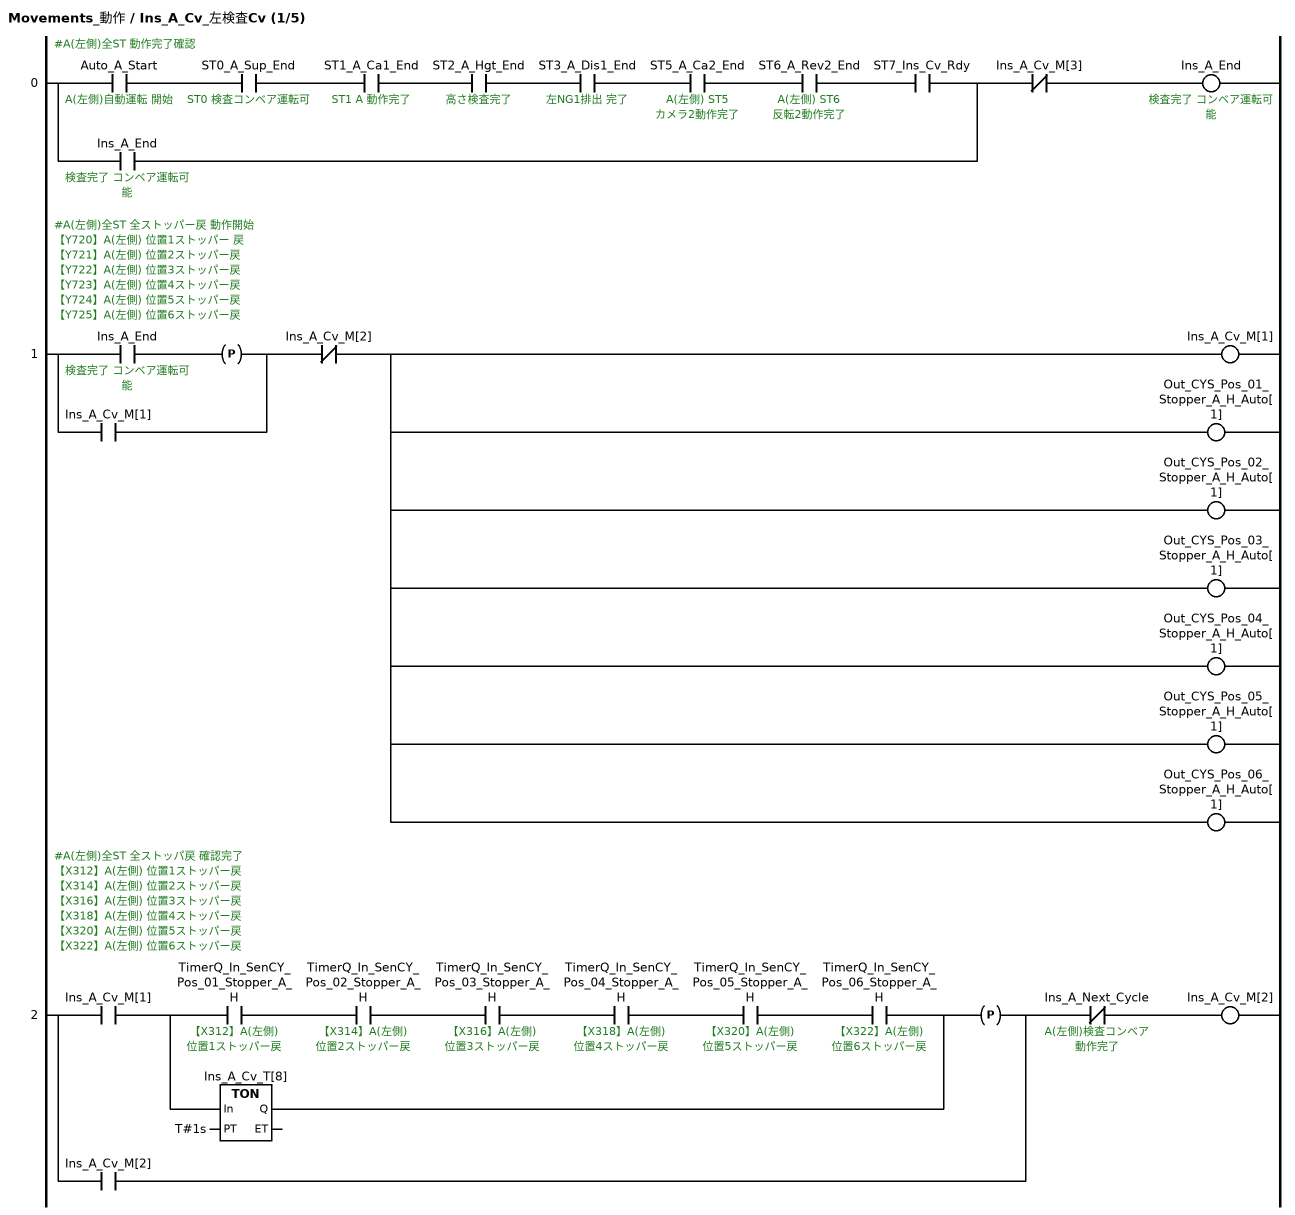
(* Rung 0: #A(左側)全ST 動作完了確認 *)
Ins_A_End := ((Auto_A_Start AND ST0_A_Sup_End AND ST1_A_Ca1_End AND ST2_A_Hgt_End AND ST3_A_Dis1_End AND ST5_A_Ca2_End AND ST6_A_Rev2_End AND ST7_Ins_Cv_Rdy) OR Ins_A_End) AND NOT Ins_A_Cv_M[3];
(* Rung 1: #A(左側)全ST 全ストッパー戻 動作開始 / 【Y720】A(左側) 位置1ストッパー 戻 / 【Y721】A(左側) 位置2ストッパー戻 / 【Y722】A(左側) 位置3ストッパー戻 / 【Y723】A(左側) 位置4ストッパー戻 / 【Y724】A(左側) 位置5ストッパー戻 / 【Y725】A(左側) 位置6ストッパー戻 *)
_e1(CLK := Ins_A_End);
_p2 := (_e1.Q OR Ins_A_Cv_M[1]) AND NOT Ins_A_Cv_M[2];
Ins_A_Cv_M[1] := _p2;
Out_CYS_Pos_01_Stopper_A_H_Auto[1] := _p2;
Out_CYS_Pos_02_Stopper_A_H_Auto[1] := _p2;
Out_CYS_Pos_03_Stopper_A_H_Auto[1] := _p2;
Out_CYS_Pos_04_Stopper_A_H_Auto[1] := _p2;
Out_CYS_Pos_05_Stopper_A_H_Auto[1] := _p2;
Out_CYS_Pos_06_Stopper_A_H_Auto[1] := _p2;
(* Rung 2: #A(左側)全ST 全ストッパ戻 確認完了 / 【X312】A(左側) 位置1ストッパー戻 / 【X314】A(左側) 位置2ストッパー戻 / 【X316】A(左側) 位置3ストッパー戻 / 【X318】A(左側) 位置4ストッパー戻 / 【X320】A(左側) 位置5ストッパー戻 / 【X322】A(左側) 位置6ストッパー戻 *)
Ins_A_Cv_T[8](In := Ins_A_Cv_M[1], PT := T#1s);
_e3(CLK := (Ins_A_Cv_M[1] AND TimerQ_In_SenCY_Pos_01_Stopper_A_H AND TimerQ_In_SenCY_Pos_02_Stopper_A_H AND TimerQ_In_SenCY_Pos_03_Stopper_A_H AND TimerQ_In_SenCY_Pos_04_Stopper_A_H AND TimerQ_In_SenCY_Pos_05_Stopper_A_H AND TimerQ_In_SenCY_Pos_06_Stopper_A_H) OR Ins_A_Cv_T[8].Q);
Ins_A_Cv_M[2] := (_e3.Q OR Ins_A_Cv_M[2]) AND NOT Ins_A_Next_Cycle;

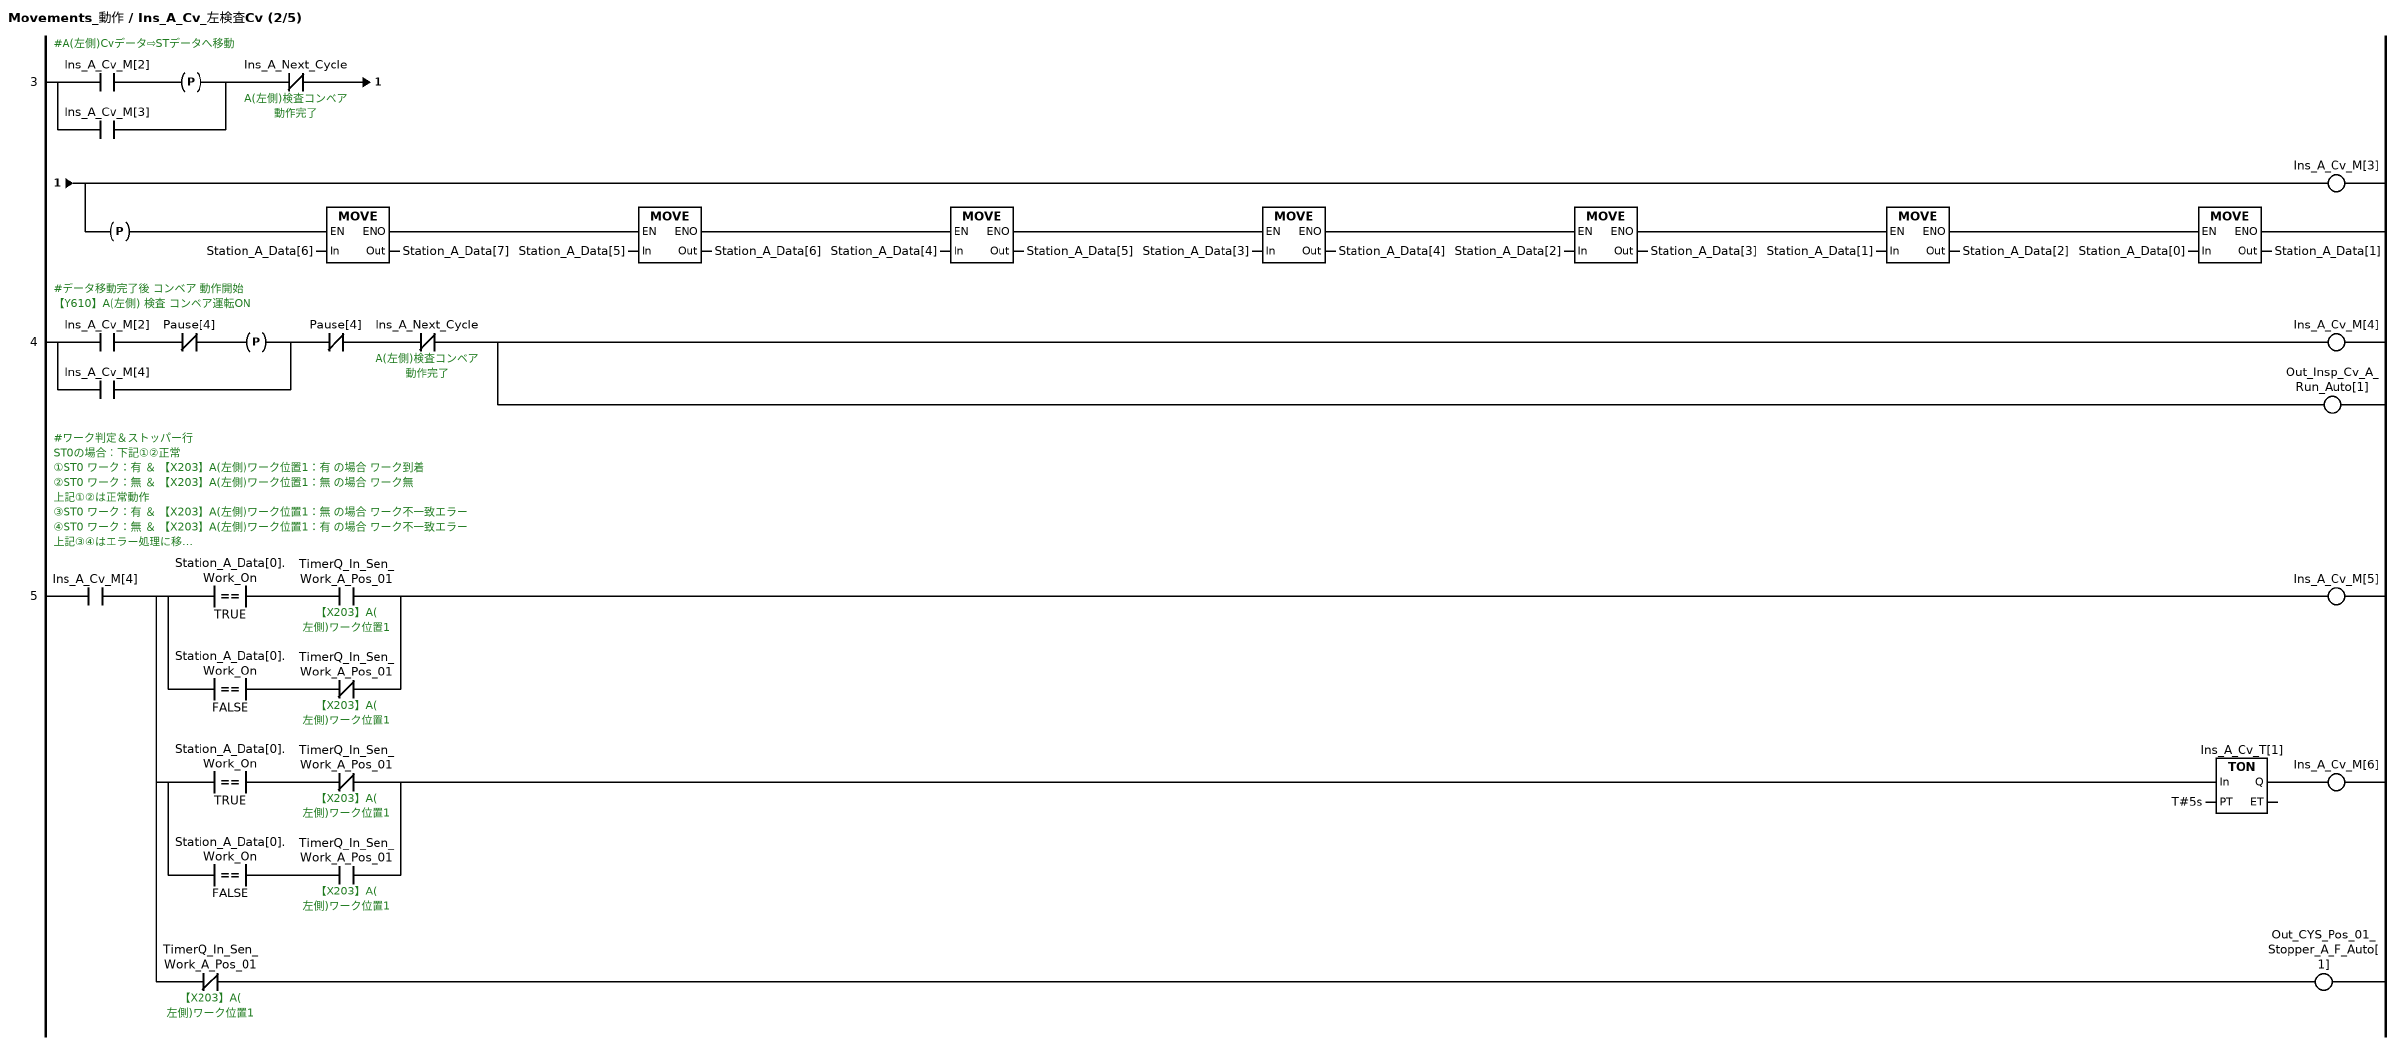
(* Rung 3: #A(左側)Cvデータ⇨STデータへ移動 *)
_e4(CLK := Ins_A_Cv_M[2]);
_p5 := (_e4.Q OR Ins_A_Cv_M[3]) AND NOT Ins_A_Next_Cycle;
Ins_A_Cv_M[3] := _p5;
_e6(CLK := _p5);
IF _e6.Q THEN
    Station_A_Data[7] := Station_A_Data[6];
    Station_A_Data[6] := Station_A_Data[5];
    Station_A_Data[5] := Station_A_Data[4];
    Station_A_Data[4] := Station_A_Data[3];
    Station_A_Data[3] := Station_A_Data[2];
    Station_A_Data[2] := Station_A_Data[1];
    Station_A_Data[1] := Station_A_Data[0];
END_IF;
(* Rung 4: #データ移動完了後 コンベア 動作開始 / 【Y610】A(左側) 検査 コンベア運転ON *)
_e7(CLK := Ins_A_Cv_M[2] AND NOT Pause[4]);
_p8 := (_e7.Q OR Ins_A_Cv_M[4]) AND NOT Pause[4] AND NOT Ins_A_Next_Cycle;
Ins_A_Cv_M[4] := _p8;
Out_Insp_Cv_A_Run_Auto[1] := _p8;
(* Rung 5: #ワーク判定＆ストッパー行 / ST0の場合：下記①②正常 / ①ST0 ワーク：有 ＆ 【X203】A(左側)ワーク位置1：有 の場合 ワーク到着 / ②ST0 ワーク：無 ＆ 【X203】A(左側)ワーク位置1：無 の場合 ワーク無 / 上記①②は正常動作 / ③ST0 ワーク：有 ＆ 【X203】A(左側)ワーク位置1：無 の場合 ワーク不一致エラー / ④ST0 ワーク：無 ＆ 【X203】A(左側)ワーク位置1：有 の場合 ワーク不一致エラー / 上記③④はエラー処理に移動 / ⑤【X203】A(左側)ワーク位置1：無 の場合 / 【Y720】A(左側) 位置1ストッパー 行 *)
_p9 := Ins_A_Cv_M[4];
Ins_A_Cv_M[5] := Ins_A_Cv_M[4] AND (((Station_A_Data[0].Work_On = TRUE) AND TimerQ_In_Sen_Work_A_Pos_01) OR ((Station_A_Data[0].Work_On = FALSE) AND NOT TimerQ_In_Sen_Work_A_Pos_01));
Ins_A_Cv_T[1](In := _p9 AND (((Station_A_Data[0].Work_On = TRUE) AND NOT TimerQ_In_Sen_Work_A_Pos_01) OR ((Station_A_Data[0].Work_On = FALSE) AND TimerQ_In_Sen_Work_A_Pos_01)), PT := T#5s);
Ins_A_Cv_M[6] := Ins_A_Cv_T[1].Q;
Out_CYS_Pos_01_Stopper_A_F_Auto[1] := _p9 AND NOT TimerQ_In_Sen_Work_A_Pos_01;

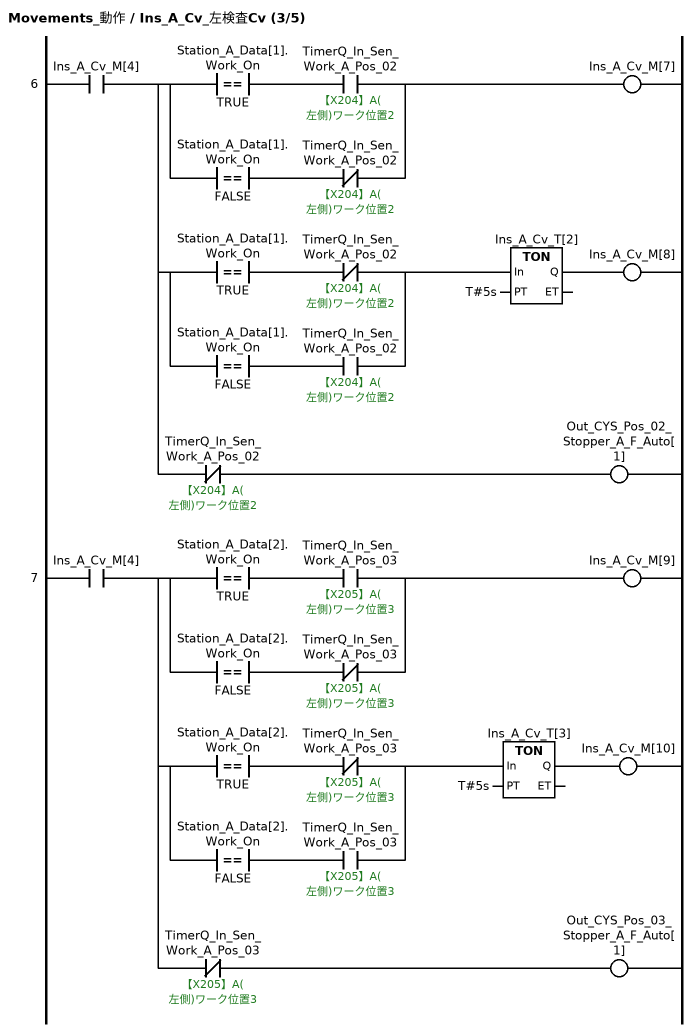
(* Rung 6 *)
_p10 := Ins_A_Cv_M[4];
Ins_A_Cv_M[7] := Ins_A_Cv_M[4] AND (((Station_A_Data[1].Work_On = TRUE) AND TimerQ_In_Sen_Work_A_Pos_02) OR ((Station_A_Data[1].Work_On = FALSE) AND NOT TimerQ_In_Sen_Work_A_Pos_02));
Ins_A_Cv_T[2](In := _p10 AND (((Station_A_Data[1].Work_On = TRUE) AND NOT TimerQ_In_Sen_Work_A_Pos_02) OR ((Station_A_Data[1].Work_On = FALSE) AND TimerQ_In_Sen_Work_A_Pos_02)), PT := T#5s);
Ins_A_Cv_M[8] := Ins_A_Cv_T[2].Q;
Out_CYS_Pos_02_Stopper_A_F_Auto[1] := _p10 AND NOT TimerQ_In_Sen_Work_A_Pos_02;
(* Rung 7 *)
_p11 := Ins_A_Cv_M[4];
Ins_A_Cv_M[9] := Ins_A_Cv_M[4] AND (((Station_A_Data[2].Work_On = TRUE) AND TimerQ_In_Sen_Work_A_Pos_03) OR ((Station_A_Data[2].Work_On = FALSE) AND NOT TimerQ_In_Sen_Work_A_Pos_03));
Ins_A_Cv_T[3](In := _p11 AND (((Station_A_Data[2].Work_On = TRUE) AND NOT TimerQ_In_Sen_Work_A_Pos_03) OR ((Station_A_Data[2].Work_On = FALSE) AND TimerQ_In_Sen_Work_A_Pos_03)), PT := T#5s);
Ins_A_Cv_M[10] := Ins_A_Cv_T[3].Q;
Out_CYS_Pos_03_Stopper_A_F_Auto[1] := _p11 AND NOT TimerQ_In_Sen_Work_A_Pos_03;

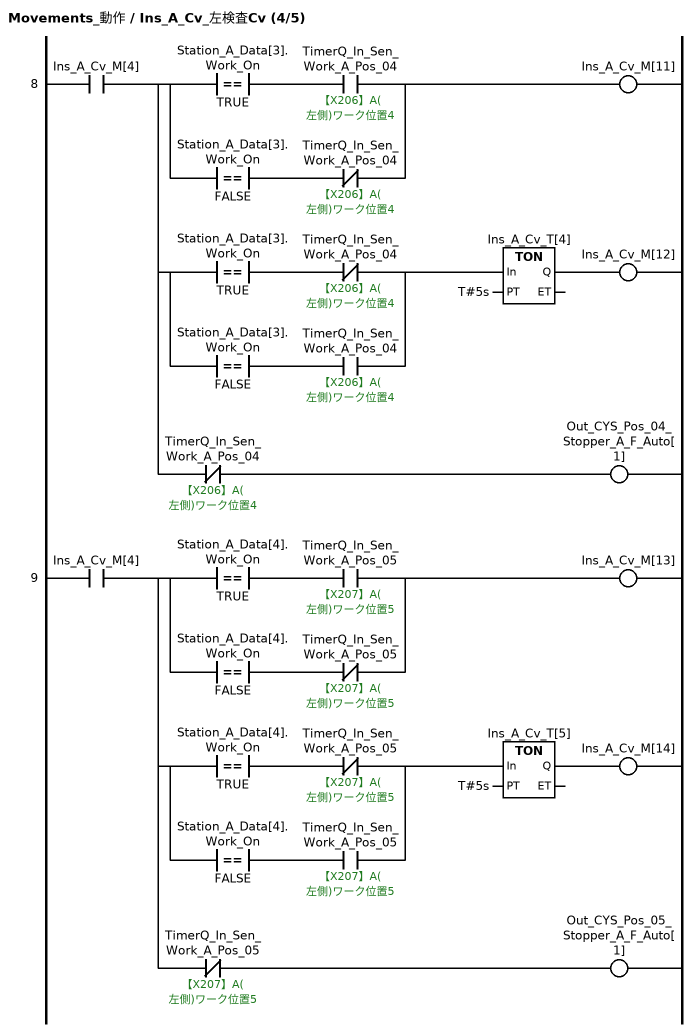
(* Rung 8 *)
_p12 := Ins_A_Cv_M[4];
Ins_A_Cv_M[11] := Ins_A_Cv_M[4] AND (((Station_A_Data[3].Work_On = TRUE) AND TimerQ_In_Sen_Work_A_Pos_04) OR ((Station_A_Data[3].Work_On = FALSE) AND NOT TimerQ_In_Sen_Work_A_Pos_04));
Ins_A_Cv_T[4](In := _p12 AND (((Station_A_Data[3].Work_On = TRUE) AND NOT TimerQ_In_Sen_Work_A_Pos_04) OR ((Station_A_Data[3].Work_On = FALSE) AND TimerQ_In_Sen_Work_A_Pos_04)), PT := T#5s);
Ins_A_Cv_M[12] := Ins_A_Cv_T[4].Q;
Out_CYS_Pos_04_Stopper_A_F_Auto[1] := _p12 AND NOT TimerQ_In_Sen_Work_A_Pos_04;
(* Rung 9 *)
_p13 := Ins_A_Cv_M[4];
Ins_A_Cv_M[13] := Ins_A_Cv_M[4] AND (((Station_A_Data[4].Work_On = TRUE) AND TimerQ_In_Sen_Work_A_Pos_05) OR ((Station_A_Data[4].Work_On = FALSE) AND NOT TimerQ_In_Sen_Work_A_Pos_05));
Ins_A_Cv_T[5](In := _p13 AND (((Station_A_Data[4].Work_On = TRUE) AND NOT TimerQ_In_Sen_Work_A_Pos_05) OR ((Station_A_Data[4].Work_On = FALSE) AND TimerQ_In_Sen_Work_A_Pos_05)), PT := T#5s);
Ins_A_Cv_M[14] := Ins_A_Cv_T[5].Q;
Out_CYS_Pos_05_Stopper_A_F_Auto[1] := _p13 AND NOT TimerQ_In_Sen_Work_A_Pos_05;

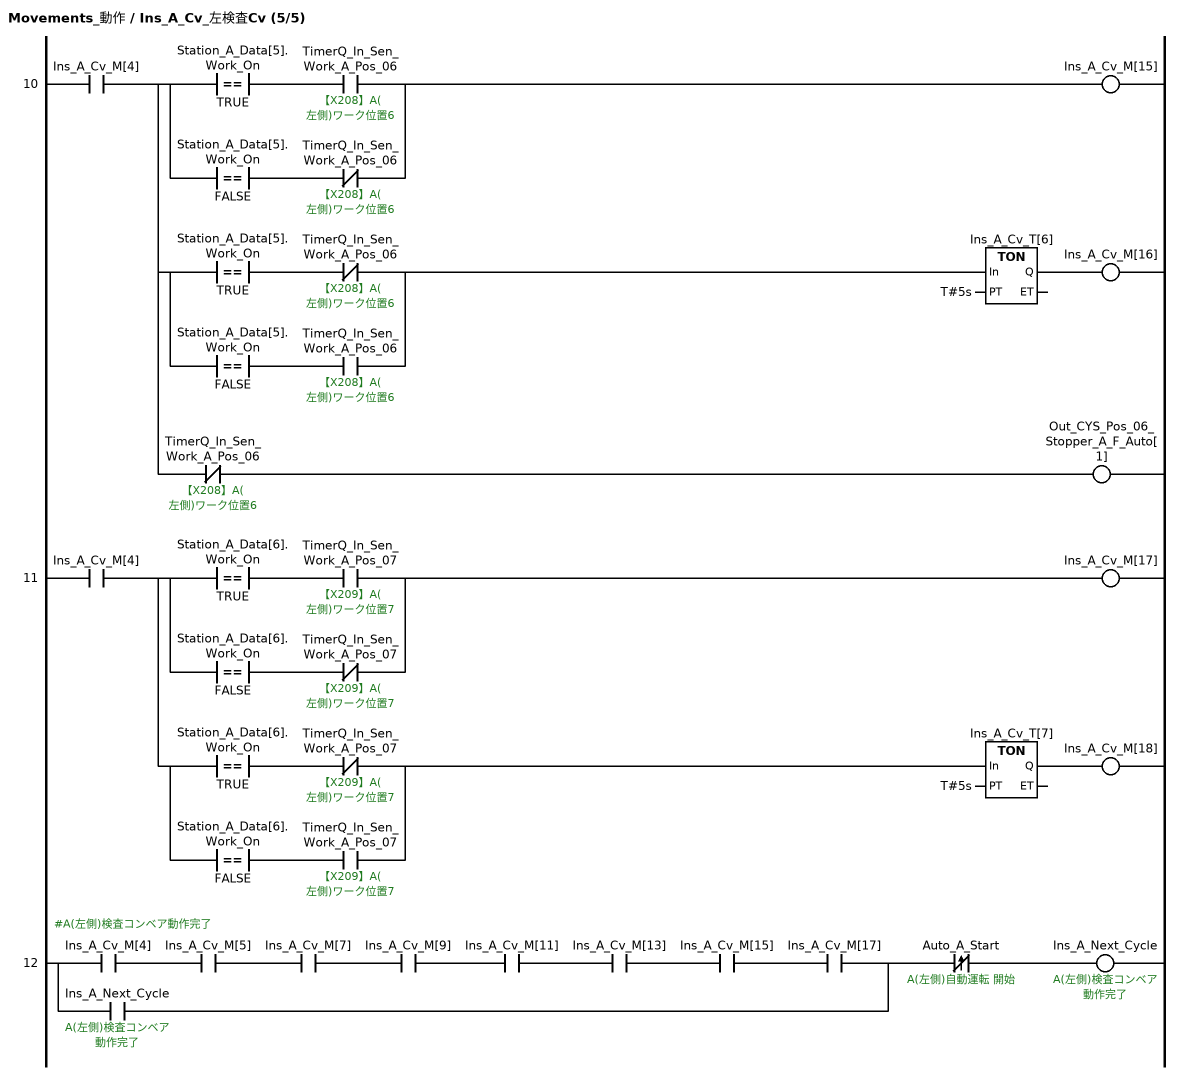
(* Rung 10 *)
_p14 := Ins_A_Cv_M[4];
Ins_A_Cv_M[15] := Ins_A_Cv_M[4] AND (((Station_A_Data[5].Work_On = TRUE) AND TimerQ_In_Sen_Work_A_Pos_06) OR ((Station_A_Data[5].Work_On = FALSE) AND NOT TimerQ_In_Sen_Work_A_Pos_06));
Ins_A_Cv_T[6](In := _p14 AND (((Station_A_Data[5].Work_On = TRUE) AND NOT TimerQ_In_Sen_Work_A_Pos_06) OR ((Station_A_Data[5].Work_On = FALSE) AND TimerQ_In_Sen_Work_A_Pos_06)), PT := T#5s);
Ins_A_Cv_M[16] := Ins_A_Cv_T[6].Q;
Out_CYS_Pos_06_Stopper_A_F_Auto[1] := _p14 AND NOT TimerQ_In_Sen_Work_A_Pos_06;
(* Rung 11 *)
_p15 := Ins_A_Cv_M[4];
Ins_A_Cv_M[17] := Ins_A_Cv_M[4] AND (((Station_A_Data[6].Work_On = TRUE) AND TimerQ_In_Sen_Work_A_Pos_07) OR ((Station_A_Data[6].Work_On = FALSE) AND NOT TimerQ_In_Sen_Work_A_Pos_07));
Ins_A_Cv_T[7](In := _p15 AND (((Station_A_Data[6].Work_On = TRUE) AND NOT TimerQ_In_Sen_Work_A_Pos_07) OR ((Station_A_Data[6].Work_On = FALSE) AND TimerQ_In_Sen_Work_A_Pos_07)), PT := T#5s);
Ins_A_Cv_M[18] := Ins_A_Cv_T[7].Q;
(* Rung 12: #A(左側)検査コンベア動作完了 *)
_e16(CLK := Auto_A_Start);
Ins_A_Next_Cycle := ((Ins_A_Cv_M[4] AND Ins_A_Cv_M[5] AND Ins_A_Cv_M[7] AND Ins_A_Cv_M[9] AND Ins_A_Cv_M[11] AND Ins_A_Cv_M[13] AND Ins_A_Cv_M[15] AND Ins_A_Cv_M[17]) OR Ins_A_Next_Cycle) AND NOT _e16.Q;

(* Section ST0_A_Sup_左供給: ladder, written here as Structured Text *)

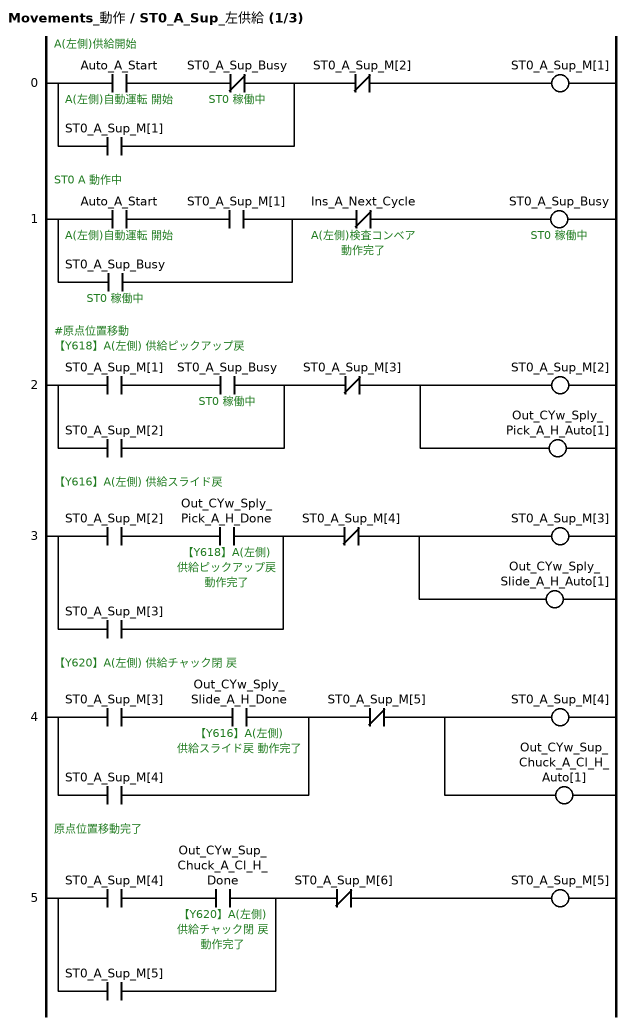
(* Rung 0: A(左側)供給開始 *)
ST0_A_Sup_M[1] := ((Auto_A_Start AND NOT ST0_A_Sup_Busy) OR ST0_A_Sup_M[1]) AND NOT ST0_A_Sup_M[2];
(* Rung 1: ST0 A 動作中 *)
ST0_A_Sup_Busy := ((Auto_A_Start AND ST0_A_Sup_M[1]) OR ST0_A_Sup_Busy) AND NOT Ins_A_Next_Cycle;
(* Rung 2: #原点位置移動 / 【Y618】A(左側) 供給ピックアップ戻 *)
_p17 := ((ST0_A_Sup_M[1] AND ST0_A_Sup_Busy) OR ST0_A_Sup_M[2]) AND NOT ST0_A_Sup_M[3];
ST0_A_Sup_M[2] := _p17;
Out_CYw_Sply_Pick_A_H_Auto[1] := _p17;
(* Rung 3: 【Y616】A(左側) 供給スライド戻 *)
_p18 := ((ST0_A_Sup_M[2] AND Out_CYw_Sply_Pick_A_H_Done) OR ST0_A_Sup_M[3]) AND NOT ST0_A_Sup_M[4];
ST0_A_Sup_M[3] := _p18;
Out_CYw_Sply_Slide_A_H_Auto[1] := _p18;
(* Rung 4: 【Y620】A(左側) 供給チャック閉 戻 *)
_p19 := ((ST0_A_Sup_M[3] AND Out_CYw_Sply_Slide_A_H_Done) OR ST0_A_Sup_M[4]) AND NOT ST0_A_Sup_M[5];
ST0_A_Sup_M[4] := _p19;
Out_CYw_Sup_Chuck_A_Cl_H_Auto[1] := _p19;
(* Rung 5: 原点位置移動完了 *)
ST0_A_Sup_M[5] := ((ST0_A_Sup_M[4] AND Out_CYw_Sup_Chuck_A_Cl_H_Done) OR ST0_A_Sup_M[5]) AND NOT ST0_A_Sup_M[6];

